//The order from Siemens is complete, nothing is remembered from earlier washes.
//Local requests of FB_CIP_Siemens carry their start too, requests of the HMI have none (item 7, 02.11.2026)
IF eReq.eClient=E_CIP_Usage.eExternal OR eReq.eStartState<>E_Element_State_Long.eOff THEN;
	eCIP_State:=eReq.eStartState;
ELSIF eReq.eType=E_CIP_Type.Full THEN;
	eCIP_State:=E_Element_State_Long.eNotClean;
ELSE;
	eCIP_State:=E_Element_State_Long.eCIP_1_Rinzed;
END_IF
g_Data.b_CIP_Run:=TRUE;
bClientRef_done:=TRUE;
END_ACTION

ACTION _aReadyToCondition_Count_active:

(*
IF TRUE 
AND pcFlow1_Rate.mRun()
AND pcFlow2_Rate.mRun()
//AND pcPressure.mRun()
THEN;
	bStepDone:=TRUE;
ELSE;
	bStepDone:=FALSE;
END_IF
*)
END_ACTION

ACTION _aReadyToCondition_Count_entry:

fb_PumpCIP.m_Run(RPM:=st_CIP_Param.r_CIP_Pump);
END_ACTION

ACTION _aReFill_Water_T93_active:
IF TRUE
//AND lvlTank_T94.e_state=E_Tank_Level.eLL
AND lvlTank_T93.rTankLevel + 0 > st_CIP_Param.r_Tank93_Volume//st_CIP_Param.r_Water_TankLvl_Lcl_1 // Client requered Level
THEN;	
	bStepDone:=TRUE;
	fbPis.m_SetByRecipe(stPis:=stPis_FillWater_T93, req:=E_Piston_Recipe_State.Release);
ELSE;
	//Fill water
	bStepDone:=FALSE;
		IF NOT arrTanksSens[E_Tank_Name.T93].get_stTankLevel_OverFlow() THEN;
			fbPis.m_SetByRecipe(stPis:=stPis_FillWater_T93, req:=E_Piston_Recipe_State.Act);			
		END_IF
END_IF
END_ACTION

ACTION _aReFill_Water_T94_active:
IF TRUE
//AND lvlTank_T94.e_state=E_Tank_Level.eLL
AND lvlTank_T94.rTankLevel +20>st_CIP_Param.r_Tank94_Volume//st_CIP_Param.r_Water_TankLvl_Lcl_1 // Client requered Level
THEN;	
	bStepDone:=TRUE;
	fbPis.m_SetByRecipe(stPis:=stPis_FillWater_T94, req:=E_Piston_Recipe_State.Release);
ELSE;
	//Fill water
	bStepDone:=FALSE;
	IF NOT arrTanksSens[E_Tank_Name.T94].get_stTankLevel_OverFlow() THEN;
		fbPis.m_SetByRecipe(stPis:=stPis_FillWater_T94, req:=E_Piston_Recipe_State.Act);			
	END_IF
END_IF
END_ACTION

ACTION _aReset_Cond_Tm_CIP2_01_active:
tonr_CIP_Condition(ResetTime:=TRUE);
END_ACTION

ACTION _aSet_Valves_ToDeafult_active:
bStepDone:=FALSE;
IF TRUE 
AND fbPis.m_CheckByRecipe(stPis:=stPis_FillWater_T91, 	req:=E_Piston_Recipe_State.Release) 
AND fbPis.m_CheckByRecipe(stPis:=stPis_FillWater_T92, 	req:=E_Piston_Recipe_State.Release) 
AND fbPis.m_CheckByRecipe(stPis:=stPis_FillWater_T93, 	req:=E_Piston_Recipe_State.Release) 
AND fbPis.m_CheckByRecipe(stPis:=stPis_FillWater_T94, 	req:=E_Piston_Recipe_State.Release) 

THEN;
	bStepDone:=TRUE;
END_IF
END_ACTION

ACTION _aSet_Valves_ToDeafult_entry:
fbPis.m_SetByRecipe(stPis:=stPis_FillWater_T91, req:=E_Piston_Recipe_State.Release);
fbPis.m_SetByRecipe(stPis:=stPis_FillWater_T92, req:=E_Piston_Recipe_State.Release);
fbPis.m_SetByRecipe(stPis:=stPis_FillWater_T93, req:=E_Piston_Recipe_State.Release);
fbPis.m_SetByRecipe(stPis:=stPis_FillWater_T94, req:=E_Piston_Recipe_State.Release);

_aDisconnect_n_Drain_CIP_Client_entry();
END_ACTION

ACTION _aSprinkler_Request_CIP1_active:


IF TRUE // Type Tank
AND bClientTypeIs_Tank	
AND bSprinkler
THEN;	
	bStepDone:=TRUE;
	m_DashState_done(stage:=E_CIP_DashStage_List.e02_CIP1_Client_Drain_Product_Rest_Sprinkler);
	
ELSIF TRUE // Type Pine
AND NOT bClientTypeIs_Tank	
THEN;	
	bStepDone:=TRUE;
	m_DashState_done(stage:=E_CIP_DashStage_List.e01_CIP1_Client_Drain_Product_Rest_Pipe);
	
ELSE;
	//continue with sprinkler
	bStepDone:=FALSE;
	m_DashState_done(stage:=E_CIP_DashStage_List.e01_CIP1_Client_Drain_Product_Rest_Pipe);
	m_DashState_activate(stage:=E_CIP_DashStage_List.e02_CIP1_Client_Drain_Product_Rest_Sprinkler);
	
END_IF
END_ACTION

ACTION _aSprinkler_Request_CIP35_active:


IF TRUE // Type Tank
AND bClientTypeIs_Tank	
AND bSprinkler
THEN;	
	bStepDone:=TRUE;
	CASE eCIP_State OF
	
		E_Element_State_Long.eCIP_2_Deterged:;
				m_DashState_done(stage:=E_CIP_DashStage_List.e11_CIP3_Detergent_Clean_Sprinkler);
	
		E_Element_State_Long.eCIP_4_Sanitized:;
				m_DashState_done(stage:=E_CIP_DashStage_List.e20_CIP5_DisInfection_Clean_Sprinkler);
				
	END_CASE	
	
ELSIF TRUE // Type Pine
AND NOT bClientTypeIs_Tank	
THEN;	
	bStepDone:=TRUE;
	CASE eCIP_State OF
	
		E_Element_State_Long.eCIP_2_Deterged:;
				m_DashState_done(stage:=E_CIP_DashStage_List.e10_CIP3_Detergent_Clean_Pipe);
	
		E_Element_State_Long.eCIP_4_Sanitized:;
				m_DashState_done(stage:=E_CIP_DashStage_List.e19_CIP5_DisInfection_Clean_Pipe);
				
	END_CASE	
	
ELSE;
	//continue with sprinkler
	bStepDone:=FALSE;
	CASE eCIP_State OF
	
		E_Element_State_Long.eCIP_2_Deterged:;
				m_DashState_done(stage:=E_CIP_DashStage_List.e10_CIP3_Detergent_Clean_Pipe);
				m_DashState_activate(stage:=E_CIP_DashStage_List.e11_CIP3_Detergent_Clean_Sprinkler);
	
		E_Element_State_Long.eCIP_4_Sanitized:;
				m_DashState_done(stage:=E_CIP_DashStage_List.e19_CIP5_DisInfection_Clean_Pipe);
				m_DashState_activate(stage:=E_CIP_DashStage_List.e20_CIP5_DisInfection_Clean_Sprinkler);
				
	END_CASE	
	
END_IF
END_ACTION

ACTION _aStartPump_CIP1_01_active:
bStepDone:=FALSE;
(*
IF StartPump_CIP1_01.t>SECOND_TO_TIME(st_CIP_Param.t_PumpInitRun) 
OR lvlTank_T93.rTankLevel<st_CIP_Param.r_Tank93_Volume//st_CIP_Param.r_RWater_93_TankLvl
THEN//Time+flow+water volume
	bStepDone:=TRUE;
END_IF
*)
bStepDone:=TRUE;
END_ACTION

ACTION _aStartPump_CIP1_01_entry:
fb_PumpCIP.m_Run(RPM:=st_CIP_Param.r_CIP_Pump);


mVolumeReset_All();

tonr_CIP_Condition(ResetTime:=TRUE);
END_ACTION

ACTION _aStartPump_CIP2_01_active:
IF TRUE 
//AND stAnalogSensor[E_ASense_Name.FT1001].Value>=g_Data.arr_CIP_Recipe[0].r_Flow_1 // 
//AND stAnalogSensor[E_ASense_Name.FT1002].Value>=g_Data.arr_CIP_Recipe[0].r_Flow_2 // 
//AND stAnalogSensor[E_ASense_Name.PT1001].Value>=g_Data.arr_CIP_Recipe[0].r_Pressure // 
//AND pcFlow1_Rate.mRun_With_SP(Set_Point:=g_Data.arr_CIP_Recipe[0].r_Flow_Pipe)
//AND pcFlow2_Rate.mRun_With_SP(Set_Point:=g_Data.arr_CIP_Recipe[0].r_Flow_Pipe)
AND pcFlow1_Rate.mRun()
AND pcFlow2_Rate.mRun()
//AND pcPressure.mRun()
THEN;
	bStepDone:=TRUE;
ELSE;
	bStepDone:=FALSE;
END_IF

fb_PumpCIP.m_Run(RPM:=pcFlow1_Rate.mRun_PID(Set_Point:=g_Data.arr_CIP_Recipe[0].r_Flow_Pipe,controlManual:=NOT(fb_PumpCIP.modeAuto)));
END_ACTION

ACTION _aStartPump_CIP2_01_entry:

//fb_PumpDetergent.m_Auto();
fb_HeatExchenger.m_Auto();
bCIP_Condition_Failed:=FALSE;
bCIP_Condition_Done:=FALSE;
iConcentrationDeluteCounter:=0;

nStepHeat:=1;
END_ACTION

ACTION _aStartPump_CIP2_02_active:
fb_PumpCIP.m_Run(RPM:=pcFlow1_Rate.mRun_PID(Set_Point:=fFlowRate, controlManual:=NOT(fb_PumpCIP.modeAuto)));


IF TRUE 
AND pcFlow1_Rate.mRun()
AND pcFlow2_Rate.mRun()
//AND pcPressure.mRun()
THEN;
	bStepDone:=TRUE;
ELSE;
	bStepDone:=FALSE;
END_IF
END_ACTION

ACTION _aStartPump_CIP2_02_entry:
fb_HeatExchenger.m_Auto();
bCIP_Condition_Failed:=FALSE;
bCIP_Condition_Done:=FALSE;
iConcentrationDeluteCounter:=0;

nStepHeat:=10;
END_ACTION

ACTION _aStartPump_CIP2_RPM_01_active:
bStepDone:=FALSE;
fb_PumpCIP.m_Run(RPM:=g_Data.arr_CIP_Recipe[0].r_CIP_Pump);//1500

IF TRUE //Future condition
AND StartPump_CIP2_RPM_01.t>SECOND_TO_TIME(g_Data.arr_CIP_Recipe[0].t_PumpInitRun) 
AND fb_PumpCIP.nRPM=g_Data.arr_CIP_Recipe[0].r_CIP_Pump
//AND stAnalogSensor[E_ASense_Name.FT1001].Value>=g_Data.arr_CIP_Recipe[0].r_Flow_Pipe // 
//AND stAnalogSensor[E_ASense_Name.FT1002].Value>=g_Data.arr_CIP_Recipe[0].r_Flow_Pipe // 
THEN;
	bStepDone:=TRUE;
END_IF
END_ACTION

ACTION _aStartPump_CIP2_RPM_02_active:
bStepDone:=FALSE;

fb_PumpCIP.m_Run(RPM:=st_CIP_Param.r_CIP_Pump);

bStepDone:=TRUE;

// to stas question ? deference:
//fb_PumpCIP.m_Run(RPM:=g_Data.arr_CIP_Recipe[0].r_CIP_Pmp_1);//1500
//fb_PumpCIP.m_Run(RPM:=st_CIP_Param.r_CIP_Pmp_1);
(*
IF TRUE //Future condition
AND delta_T92_Volume < - st_CIP_Param.r_Volume_Solution_Fill // Volume 
//AND StartPump_CIP2_RPM_02.t>SECOND_TO_TIME(g_Data.arr_CIP_Recipe[0].t_PumpInitRun) 
THEN;
	bStepDone:=TRUE;
END_IF
*)
END_ACTION

ACTION _aStartPump_CIP2_RPM_02_entry:
mVolumeReset_All();
tonr_CIP_Condition(ResetTime:=TRUE);
END_ACTION

ACTION _aStartPump_CIP4_RPM_01_active:
bStepDone:=FALSE;
fb_PumpCIP.m_Run(RPM:=g_Data.arr_CIP_Recipe[0].r_CIP_Pump);

IF TRUE //Future condition
AND StartPump_CIP4_RPM_01.t>SECOND_TO_TIME(g_Data.arr_CIP_Recipe[0].t_PumpInitRun) 
THEN;
	bStepDone:=TRUE;
END_IF
END_ACTION

ACTION _aStartPump_CIP4_RPM_02_active:
bStepDone:=FALSE;
fb_PumpCIP.m_Run(RPM:=pcFlow1_Rate.mRun_PID(Set_Point:=st_CIP_Param.r_CIP_Pump,controlManual:=NOT(fb_PumpCIP.modeAuto)));


IF TRUE //Future condition
AND StartPump_CIP4_RPM_02.t>SECOND_TO_TIME(st_CIP_Param.t_PumpInitRun) 
THEN;
	bStepDone:=TRUE;
END_IF
END_ACTION

ACTION _aStartPump_CIP4_01_active:
IF TRUE 
(*AND stAnalogSensor[E_ASense_Name.FT1001].Value>=g_Data.arr_CIP_Recipe[0].r_Flow_1//200 // 
AND stAnalogSensor[E_ASense_Name.FT1002].Value>=g_Data.arr_CIP_Recipe[0].r_Flow_2//200 // 
AND stAnalogSensor[E_ASense_Name.PT1001].Value>=g_Data.arr_CIP_Recipe[0].r_Pressure//0.5 //*)
AND pcFlow1_Rate.mRun()
AND pcFlow2_Rate.mRun()
//AND pcPressure.mRun()
THEN;
	bStepDone:=TRUE;
ELSE;
	bStepDone:=FALSE;
END_IF

fb_PumpCIP.m_Run(RPM:=pcFlow1_Rate.mRun_PID(Set_Point:=g_Data.arr_CIP_Recipe[0].r_Flow_Pipe,controlManual:=NOT(fb_PumpCIP.modeAuto)));
END_ACTION

ACTION _aStartPump_CIP4_01_entry:


fb_HeatExchenger.m_Auto();
bCIP_Condition_Failed:=FALSE;
bCIP_Condition_Done:=FALSE;

nStepHeat:=2;
iConcentrationDeluteCounter:=0;
END_ACTION

ACTION _aStartPump_CIP4_02_active:
IF TRUE 
(*AND stAnalogSensor[E_ASense_Name.FT1001].Value>=st_CIP_Param.r_Flow_1 // 
AND stAnalogSensor[E_ASense_Name.FT1002].Value>=st_CIP_Param.r_Flow_2 // 
AND stAnalogSensor[E_ASense_Name.PT1001].Value>=st_CIP_Param.r_Pressure // *)
AND pcFlow1_Rate.mRun()
AND pcFlow2_Rate.mRun()
//AND pcPressure.mRun()
THEN;
	bStepDone:=TRUE;
ELSE;
	bStepDone:=FALSE;
END_IF

//fb_PumpCIP.m_Run(RPM:=pcFlow1_Rate.mRun_PID(Set_Point:=fFlowRate,controlManual:=NOT(fb_PumpCIP.modeAuto)));

IF TRUE //Future condition
AND StartPump_CIP4_02.t>SECOND_TO_TIME(st_CIP_Param.t_PumpInitRun) THEN;
	fb_PumpCIP.m_Run(RPM:=pcFlow1_Rate.mRun_PID(Set_Point:=fFlowRate,controlManual:=NOT(fb_PumpCIP.modeAuto)));
	
END_IF

IF NOT bSprinkler THEN
	//pipe
	tConditionTime	:=st_CIP_Param.t_ConditionDisInfection;
	fFlowRate		:=st_CIP_Param.r_Flow_Pipe;
	//rVolume_Collect :=st_CIP_Param.r_Volume_Collect_DisInfection;
	//rVolume_Drain	:=st_CIP_Param.r_Volume_Drain_DisInfection;
	//rVolume_Recycle	:=st_CIP_Param.r_Volume_Recycle_DisInfection;
ELSE
	//sprinkler
	tConditionTime	:=st_CIP_Param.t_ConditionDisInfection_Sprinkler;
	fFlowRate		:=st_CIP_Param.r_Flow_Sprinkler;
	//rVolume_Collect :=st_CIP_Param.r_Volume_Collect_DisInfection*st_CIP_Param.r_Volume_Sprinkler_Ratio;
	//rVolume_Drain	:=st_CIP_Param.r_Volume_Drain_DisInfection*st_CIP_Param.r_Volume_Sprinkler_Ratio;
	//rVolume_Recycle	:=st_CIP_Param.r_Volume_Recycle_DisInfection*st_CIP_Param.r_Volume_Sprinkler_Ratio;
END_IF
END_ACTION

ACTION _aStartPump_CIP4_02_entry:

//fb_PumpDisinfection.m_Auto();
	
//Heat Exchenger	
fb_HeatExchenger.m_Auto();

bCIP_Condition_Failed:=FALSE;
bCIP_Condition_Done:=FALSE;
iConcentrationDeluteCounter:=0;

nStepHeat:=20;
END_ACTION

ACTION _aStartPump_CIP35_active:
bStepDone:=FALSE;
IF TRUE 
//AND fbPis.m_CheckByRecipe(stPis:=stPis_FillWater_T94, 		req:=E_Piston_Recipe_State.NoChanges) 
THEN
	//bStepDone:=TRUE;
END_IF
bStepDone:=TRUE;
END_ACTION

ACTION _aStartPump_CIP35_entry:
//fbPis.m_SetByRecipe(stPis:=stPis_FillWater_T94, 	req:=E_Piston_Recipe_State.NoChanges);
fb_PumpCIP.m_Run(RPM:=st_CIP_Param.r_CIP_Pump);


mVolumeReset_All();
bSprinkler:=FALSE;
tonr_CIP_Condition(ResetTime:=TRUE);
END_ACTION

ACTION _aStop_Pump_entry:
fb_PumpCIP.m_Stop();


fb_PumpDetergent.m_Stop();
fb_PumpDisinfection.m_Stop();
END_ACTION

ACTION _aStopPump_CIP1_01_entry:
fb_PumpCIP.m_Stop();
END_ACTION

ACTION _aStopPump_CIP1_02_entry:
fb_PumpCIP.m_Stop();
END_ACTION

ACTION _aStopPump_CIP2_01_entry:
fb_PumpCIP.m_Stop();

m_DashState_done(stage:=E_CIP_DashStage_List.e04_CIP2_Local_Detergent_Condition);
END_ACTION

ACTION _aStopPump_CIP2_02_entry:
fb_PumpCIP.m_Stop();
END_ACTION

ACTION _aStopPump_CIP2_03_entry:
fb_PumpCIP.m_Stop();
END_ACTION

ACTION _aStopPump_CIP4_01_entry:
fb_PumpCIP.m_Stop();

m_DashState_done(stage:=E_CIP_DashStage_List.e13_CIP4_Local_DisInfection_Condition);
END_ACTION

ACTION _aStopPump_CIP4_02_entry:
fb_PumpCIP.m_Stop();
END_ACTION

ACTION _aStopPump_CIP4_03_entry:
fb_PumpCIP.m_Stop();
END_ACTION

ACTION _aStopPump_CIP35_01_entry:
fb_PumpCIP.m_Stop();
END_ACTION

ACTION _aStopPump_CIP35_02_entry:
fb_PumpCIP.m_Stop();
END_ACTION

ACTION _aTank_LowLevel_CIP1_01_active:
bStepDone:=m_Check_ProductionTank_Low_Level();
END_ACTION

ACTION _aTank_LowLevel_CIP1_02_active:
bStepDone:=m_Check_ProductionTank_Low_Level();
END_ACTION

ACTION _aTank_LowLevel_CIP1_02_entry:
fb_PumpCIP.m_Stop();
END_ACTION

ACTION _aTank_LowLevel_CIP2_01_active:
bStepDone:=m_Check_ProductionTank_Low_Level();
END_ACTION

ACTION _aTank_LowLevel_CIP2_02_active:
bStepDone:=m_Check_ProductionTank_Low_Level();
END_ACTION

ACTION _aTank_LowLevel_CIP2_02_entry:
fb_PumpCIP.m_Stop();
END_ACTION

ACTION _aTank_LowLevel_CIP4_01_active:
bStepDone:=m_Check_ProductionTank_Low_Level();
END_ACTION

ACTION _aTank_LowLevel_CIP4_02_active:
bStepDone:=m_Check_ProductionTank_Low_Level();
END_ACTION

ACTION _aTank_LowLevel_CIP4_02_entry:
fb_PumpCIP.m_Stop();
END_ACTION

ACTION _aTank_LowLevel_CIP35_01_active:
bStepDone:=m_Check_ProductionTank_Low_Level();
END_ACTION

ACTION _aTank_LowLevel_CIP35_02_active:
bStepDone:=m_Check_ProductionTank_Low_Level();
END_ACTION

ACTION _aTank_LowLevel_CIP35_02_entry:
fb_PumpCIP.m_Stop();
END_ACTION

ACTION _aTank_MixProof_Clean_CIP2_active:
//Mix-proof valves are on the plant side
bStepDone:=TRUE;
END_ACTION

ACTION _aTank_MixProof_Clean_CIP2_entry:
fb_PumpCIP.m_Stop();
END_ACTION

ACTION _aTank_MixProof_Clean_CIP4_active:
//Mix-proof valves are on the plant side
bStepDone:=TRUE;
END_ACTION

ACTION _aTank_MixProof_Clean_CIP4_entry:
fb_PumpCIP.m_Stop();
END_ACTION

ACTION _aTriBlender_Selection_active:
bStepDone:=TRUE;
END_ACTION

ACTION _aTriBlender_Selection_entry:

END_ACTION

ACTION _aWaiting_Client_Drain_Done_active:
// The command from Set_Valves_ToDeafult is lost if a sub-FB was in Init or busy: give it again
IF fbCIP_Source.m_IsFree() AND NOT fbCIP_Source.m_CheckStatus(eReqStatus:=E_CIP_Source.eClose) THEN;
	fbCIP_Source.m_Run(eReqProc:=E_CIP_Source.eClose);
END_IF
IF fbCIP_Usage.m_IsFree() AND NOT fbCIP_Usage.m_CheckStatus(eReqStatus:=E_CIP_Usage.eLocal) THEN;
	fbCIP_Usage.m_Run(eReqProc:=E_CIP_Usage.eLocal);
END_IF
IF fbCIP_Return.m_IsFree() AND NOT fbCIP_Return.m_CheckStatus(eReqStatus:=E_CIP_Return.eDrain) THEN;
	fbCIP_Return.m_Run(eReqProc:=E_CIP_Return.eDrain);
END_IF

_aDisconnect_n_Drain_CIP_Client_active();
END_ACTION

ACTION act_CallProcessControl:
//Heat Exchanger
	stHeatExchanger.rValue:=g_AnalogSensor.stAnalogSensor[E_ASense_Name.TT1105].Value;
	//stHeatExchanger.rSetPoint:=st_CIP_Param.r_Temper_ClientReturn;
	pcHeatExchanger(stProcessControl:=stHeatExchanger );
//Client temperature return
	stTemp_ClntReturn.rValue:=g_AnalogSensor.stAnalogSensor[E_ASense_Name.TT1101].Value;//gIO.fbScaleFactor[E_ASense_Name.TT1101].rValOut;
	//stTemp_ClntReturn.rSetPoint:=st_CIP_Param.n _ClientReturn;
	pcTemp_ClntReturn(stProcessControl:=stTemp_ClntReturn );

//Detergent
	//Concentration
	stDetergent.rValue:=g_AnalogSensor.stAnalogSensor[E_ASense_Name.CT1101_3].Value;
	//###stDetergent.ToleranceHigh:=0.05;
	//###stDetergent.ToleravceLow:=0.05;
	//###stDetergent.rSetPoint:=st_CIP_Param.r_DetergentConcentration;//0.3;
	pcDetergent(stProcessControl:=stDetergent );
		
	//Temperature
	//stTemperature_Deterg.rValue:=testTemperature;
	stTemperature_Deterg.rValue:=g_AnalogSensor.stAnalogSensor[E_ASense_Name.TT1003].Value;
	//###stTemperature_Deterg.ToleranceHigh:=1;
	//###stTemperature_Deterg.ToleravceLow:=1;
	//###stTemperature_Deterg.rSetPoint:=st_CIP_Param.r_Temper_Detergent;
	pcTemperature_Deterg(stProcessControl:=stTemperature_Deterg );


//Disinfectant
	//Concentration
	stDisInfectant.rValue:=g_AnalogSensor.stAnalogSensor[E_ASense_Name.CT1101_4].Value;
	//###stDisInfectant.ToleranceHigh:=0.05;
	//###stDisInfectant.ToleravceLow:=0.05;
	//###stDisInfectant.rSetPoint:=st_CIP_Param.r_DisInfectionConcentration;//0.3;
	pcDisInfectant(stProcessControl:=stDisInfectant );
		
	//Temperature	
	//stTemperature_Dis.rValue:=testTemperature;
	stTemperature_Dis.rValue:=g_AnalogSensor.stAnalogSensor[E_ASense_Name.TT1004].Value;
	//###stTemperature_Dis.ToleranceHigh:=1;//0.5
	//###stTemperature_Dis.ToleravceLow:=1;//0.5
	//###stTemperature_Dis.rSetPoint:=st_CIP_Param.r_Temper_DisInfection;//65;
	pcTemperature_Dis(stProcessControl:=stTemperature_Dis );	
	
// Flow_Rate
	//CIP Pump
		//Pump CIP infeed
		stFlow1_Rate.rValue:=g_AnalogSensor.stAnalogSensor[E_ASense_Name.FT1001].Value;
		stFlow1_Rate.rValue:=g_AnalogSensor.stAnalogSensor[E_ASense_Name.FT1001].Value;
		stFlow1_Rate.rValue_Min_To_ReleaseControl:=50;// Litter/Hours
		//stFlow1_Rate.rSetPoint:=st_CIP_Param.r_Flow_Pipe;//:=150
		stFlow1_Rate.bPause:=stOper[E_ModeZone.eCIP].iActOperation=E_OperationButtons.ePauseAll;
		stFlow1_Rate.fCtrlOutput_Manual:=fb_PumpCIP.nRPM;
		stFlow1_Rate.fCtrlOutput_Max:=1700;
		stFlow1_Rate.fCtrlOutput_Min:=700;
		pcFlow1_Rate(stProcessControl:=stFlow1_Rate, );

		//Pump CIP return 
		stFlow2_Rate.rValue:=g_AnalogSensor.stAnalogSensor[E_ASense_Name.FT1002].Value;
		stFlow3_Rate.rValue:=g_AnalogSensor.stAnalogSensor[E_ASense_Name.FT1002].Value;
		stFlow3_Rate.rSetPoint:=stFlow2_Rate.rSetPoint;
		pcFlow2_Rate(stProcessControl:=stFlow2_Rate );
		pcFlow3_Rate(stProcessControl:=stFlow3_Rate );

		// TBD : to check if the first loop(local prepare) when Client selected gets relevant Flow SetPoint 
		IF bSprinkler THEN
			stFlow1_Rate.rSetPoint:=st_CIP_Param.r_Flow_Sprinkler;
			stFlow2_Rate.rSetPoint:=st_CIP_Param.r_Flow_Sprinkler;
		ELSE
			stFlow1_Rate.rSetPoint:=st_CIP_Param.r_Flow_Pipe;
			stFlow2_Rate.rSetPoint:=st_CIP_Param.r_Flow_Pipe;
		END_IF		
		
	//CIP Client Color pump
		//stFlow_Rate.rSetPoint:=150;
	//CIP Client Marinada pump
		//stFlow_Rate.rSetPoint:=150;
		
//Presure
		stP1001_Pressure.rValue:=g_AnalogSensor.stAnalogSensor[E_ASense_Name.PT1001].Value;
		pcP1001_Pressure(stProcessControl:=stP1001_Pressure );


//Load def set points
IF bLoadDefSetPoints THEN
	bLoadDefSetPoints:=FALSE;
	mLoadDefProcessSetPoints();
END_IF
		
//selecting set point based on user
	
	IF bTestPID THEN;
		pcFlow1_Rate.mRun();

		fb_PumpCIP.m_Auto(control:=pcFlow1_Rate.mRun_PID(Set_Point:=180,controlManual:=NOT(fb_PumpCIP.modeAuto)));
		
		//by CIP Pump RPM control		
		
		IF fb_PumpCIP.modeAuto THEN;
			stFlow1_Rate.bManual:=FALSE;
		ELSE;
			stFlow1_Rate.bManual:=TRUE;
			stFlow1_Rate.fCtrlOutput_Manual:=fb_PumpCIP.nRPM;
		END_IF
		
			
	END_IF
END_ACTION

ACTION act_GetReference:
stPis_FillWater_T91 REF= stPis[valFillWater_T91];
stPis_FillWater_T92 REF= stPis[valFillWater_T92];
stPis_FillWater_T93 REF= stPis[valFillWater_T93];
stPis_FillWater_T94 REF= stPis[valFillWater_T94];

	//concentration
stDetergent 	REF=g_ProcControl.arr_stProcCntrl[E_ProcessControl_Name.eDetergentConc];
pcDetergent 	REF=g_ProcControl.arr_fbProcCntrl[E_ProcessControl_Name.eDetergentConc];

stDisInfectant 	REF=g_ProcControl.arr_stProcCntrl[E_ProcessControl_Name.eDisinfectionConc];
pcDisInfectant 	REF=g_ProcControl.arr_fbProcCntrl[E_ProcessControl_Name.eDisinfectionConc];

	//Temperature
stTemperature_Deterg REF=g_ProcControl.arr_stProcCntrl[E_ProcessControl_Name.eDeterTemp];
pcTemperature_Deterg REF=g_ProcControl.arr_fbProcCntrl[E_ProcessControl_Name.eDeterTemp];

stTemperature_Dis 	 REF=g_ProcControl.arr_stProcCntrl[E_ProcessControl_Name.eDisTemp];
pcTemperature_Dis 	 REF=g_ProcControl.arr_fbProcCntrl[E_ProcessControl_Name.eDisTemp];
	//Flow rate
stFlow1_Rate REF=g_ProcControl.arr_stProcCntrl[E_ProcessControl_Name.eCIP_Flow_1];
pcFlow1_Rate REF=g_ProcControl.arr_fbProcCntrl[E_ProcessControl_Name.eCIP_Flow_1];

stFlow2_Rate REF=g_ProcControl.arr_stProcCntrl[E_ProcessControl_Name.eCIP_Flow_2];
pcFlow2_Rate REF=g_ProcControl.arr_fbProcCntrl[E_ProcessControl_Name.eCIP_Flow_2];

stFlow3_Rate REF=g_ProcControl.arr_stProcCntrl[E_ProcessControl_Name.eCIP_Flow_3];
pcFlow3_Rate REF=g_ProcControl.arr_fbProcCntrl[E_ProcessControl_Name.eCIP_Flow_3];

	//Level

	//Pressure
stP1001_Pressure 	REF=g_ProcControl.arr_stProcCntrl[E_ProcessControl_Name.eCIP_Pressure];
pcP1001_Pressure 	REF=g_ProcControl.arr_fbProcCntrl[E_ProcessControl_Name.eCIP_Pressure];

//temperature control
stTemp_ClntReturn REF=g_ProcControl.arr_stProcCntrl[E_ProcessControl_Name.eClientReturn_Temp];
pcTemp_ClntReturn REF=g_ProcControl.arr_fbProcCntrl[E_ProcessControl_Name.eClientReturn_Temp];

stHeatExchanger REF=g_ProcControl.arr_stProcCntrl[E_ProcessControl_Name.eHeatExchanger];
pcHeatExchanger REF=g_ProcControl.arr_fbProcCntrl[E_ProcessControl_Name.eHeatExchanger];
END_ACTION

ACTION act_HeatExchng:
//calling heat exchanger 
fb_HeatExchenger(stHeatExchanger:=g_Data.stHeatExchanger );

//Choosing heat exchanger set point 

CASE nStepHeat OF
	0:	
	(*	//heat excahnger not in use 
	1:
		//detergent local
		IF stTemperature_Deterg.Control_ON THEN
			g_Data.stHeatExchanger:=stTemperature_Deterg.Control_Value;
		ELSE
			g_Data.stHeatExchanger:=0;
		END_IF
	10:
		//detergent client
	2:
		//disinfection
		IF stTemperature_Dis.Control_ON THEN
			g_Data.stHeatExchanger:=stTemperature_Dis.Control_Value;
		ELSE
			g_Data.stHeatExchanger:=0;
		END_IF
	20:
		//disinfection client
	3:
		//something else
		*)
END_CASE
END_ACTION

ACTION act_Oper:
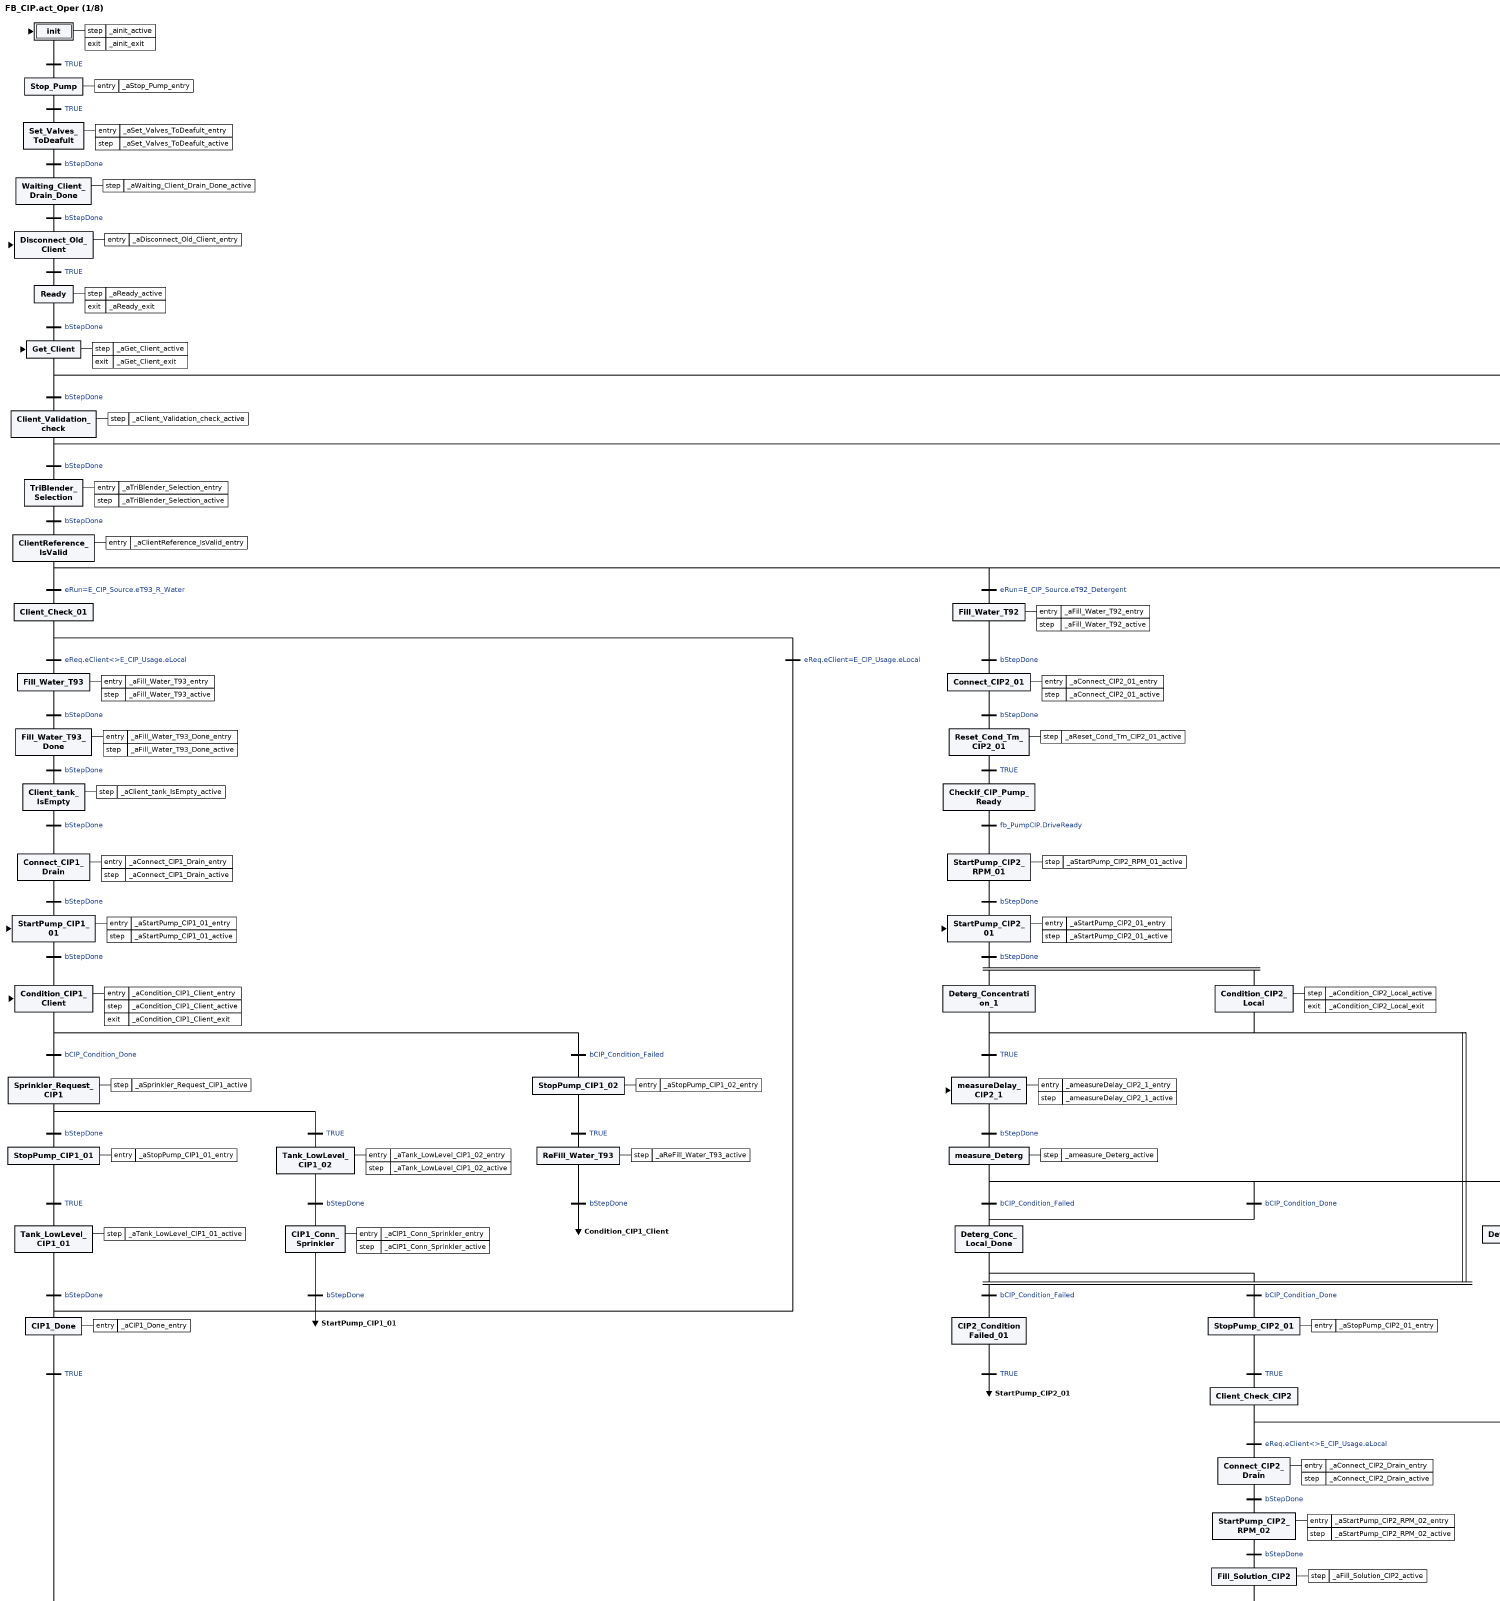
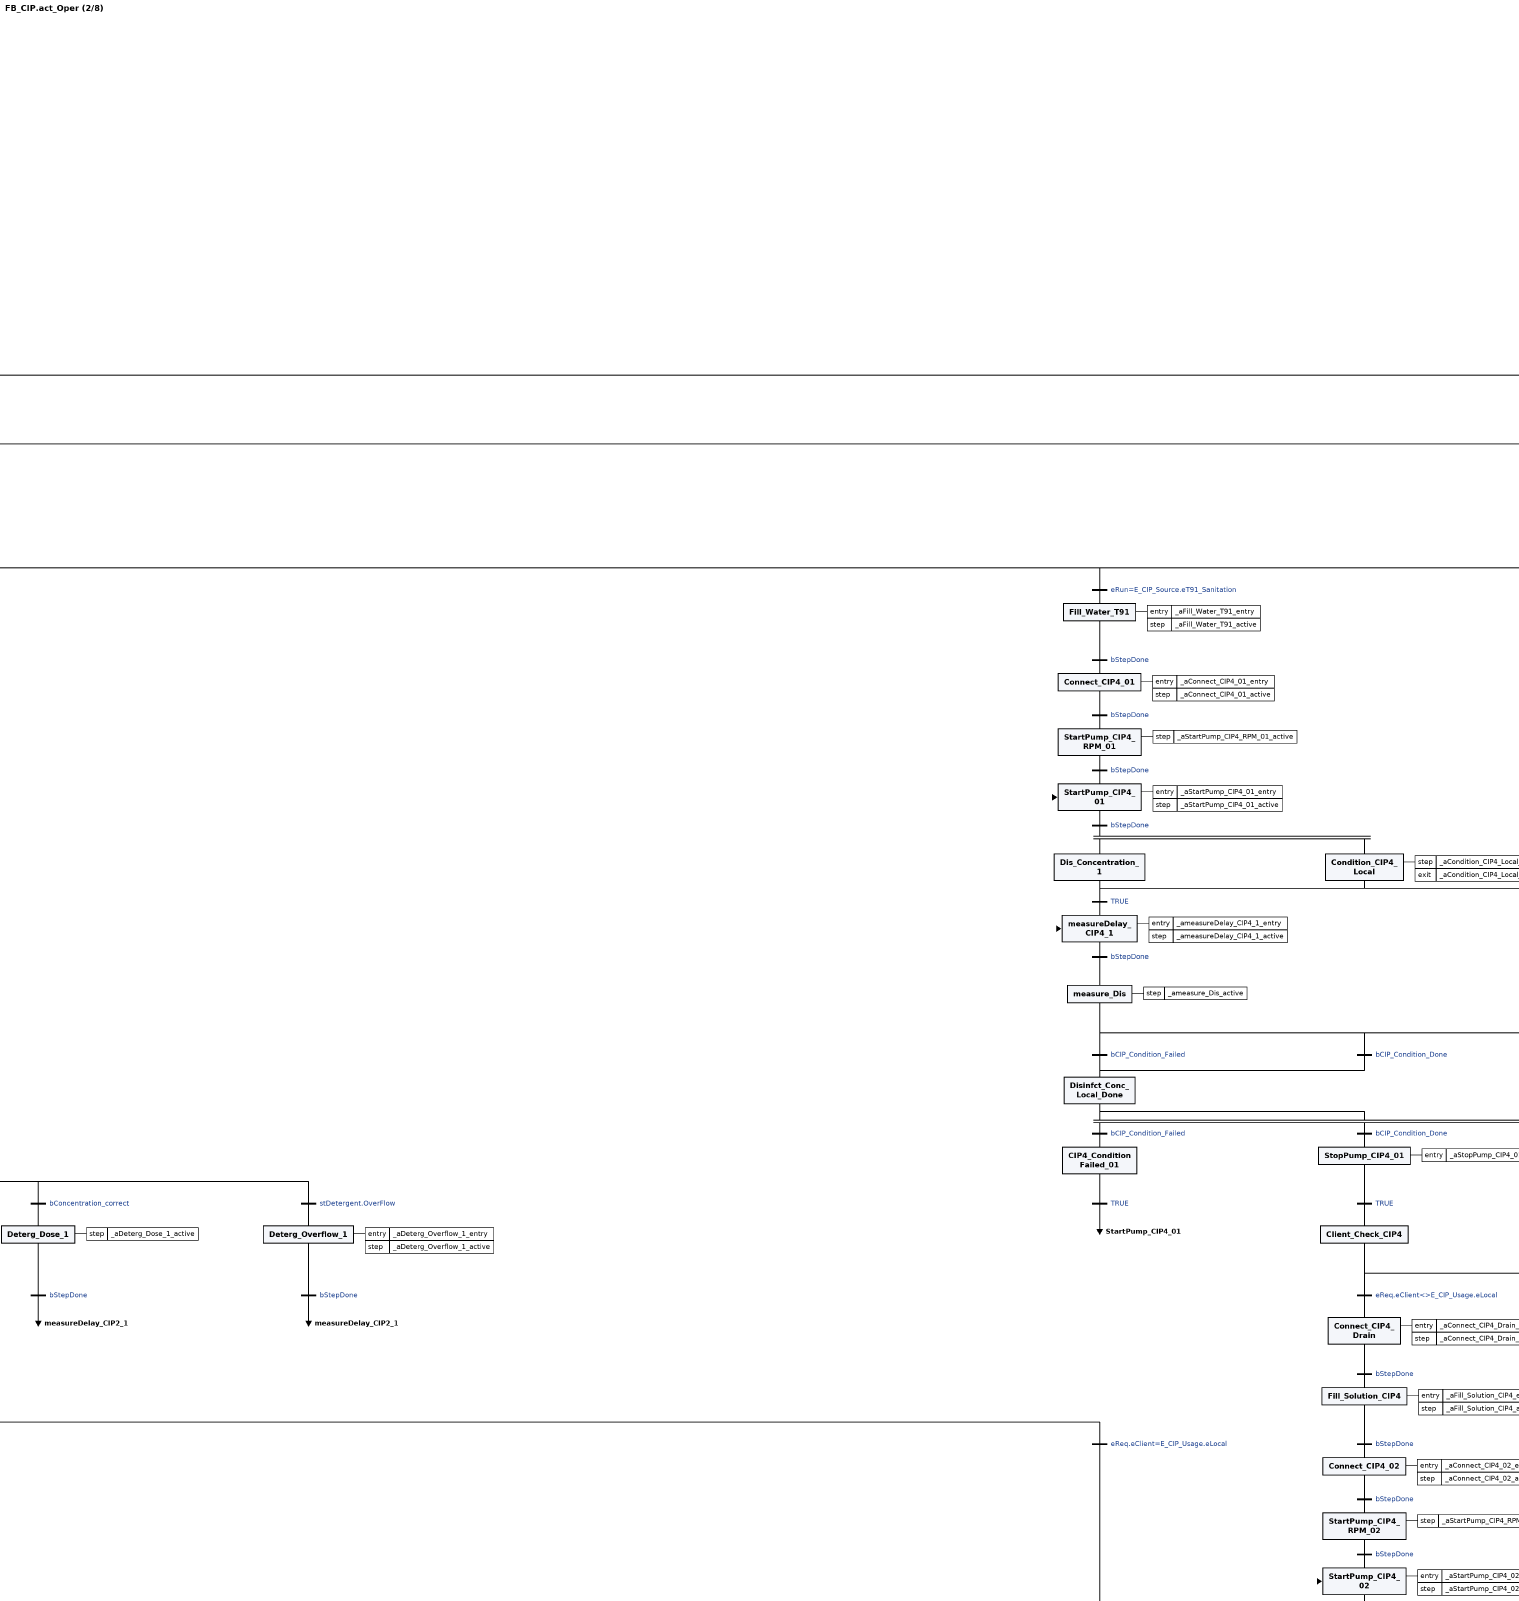
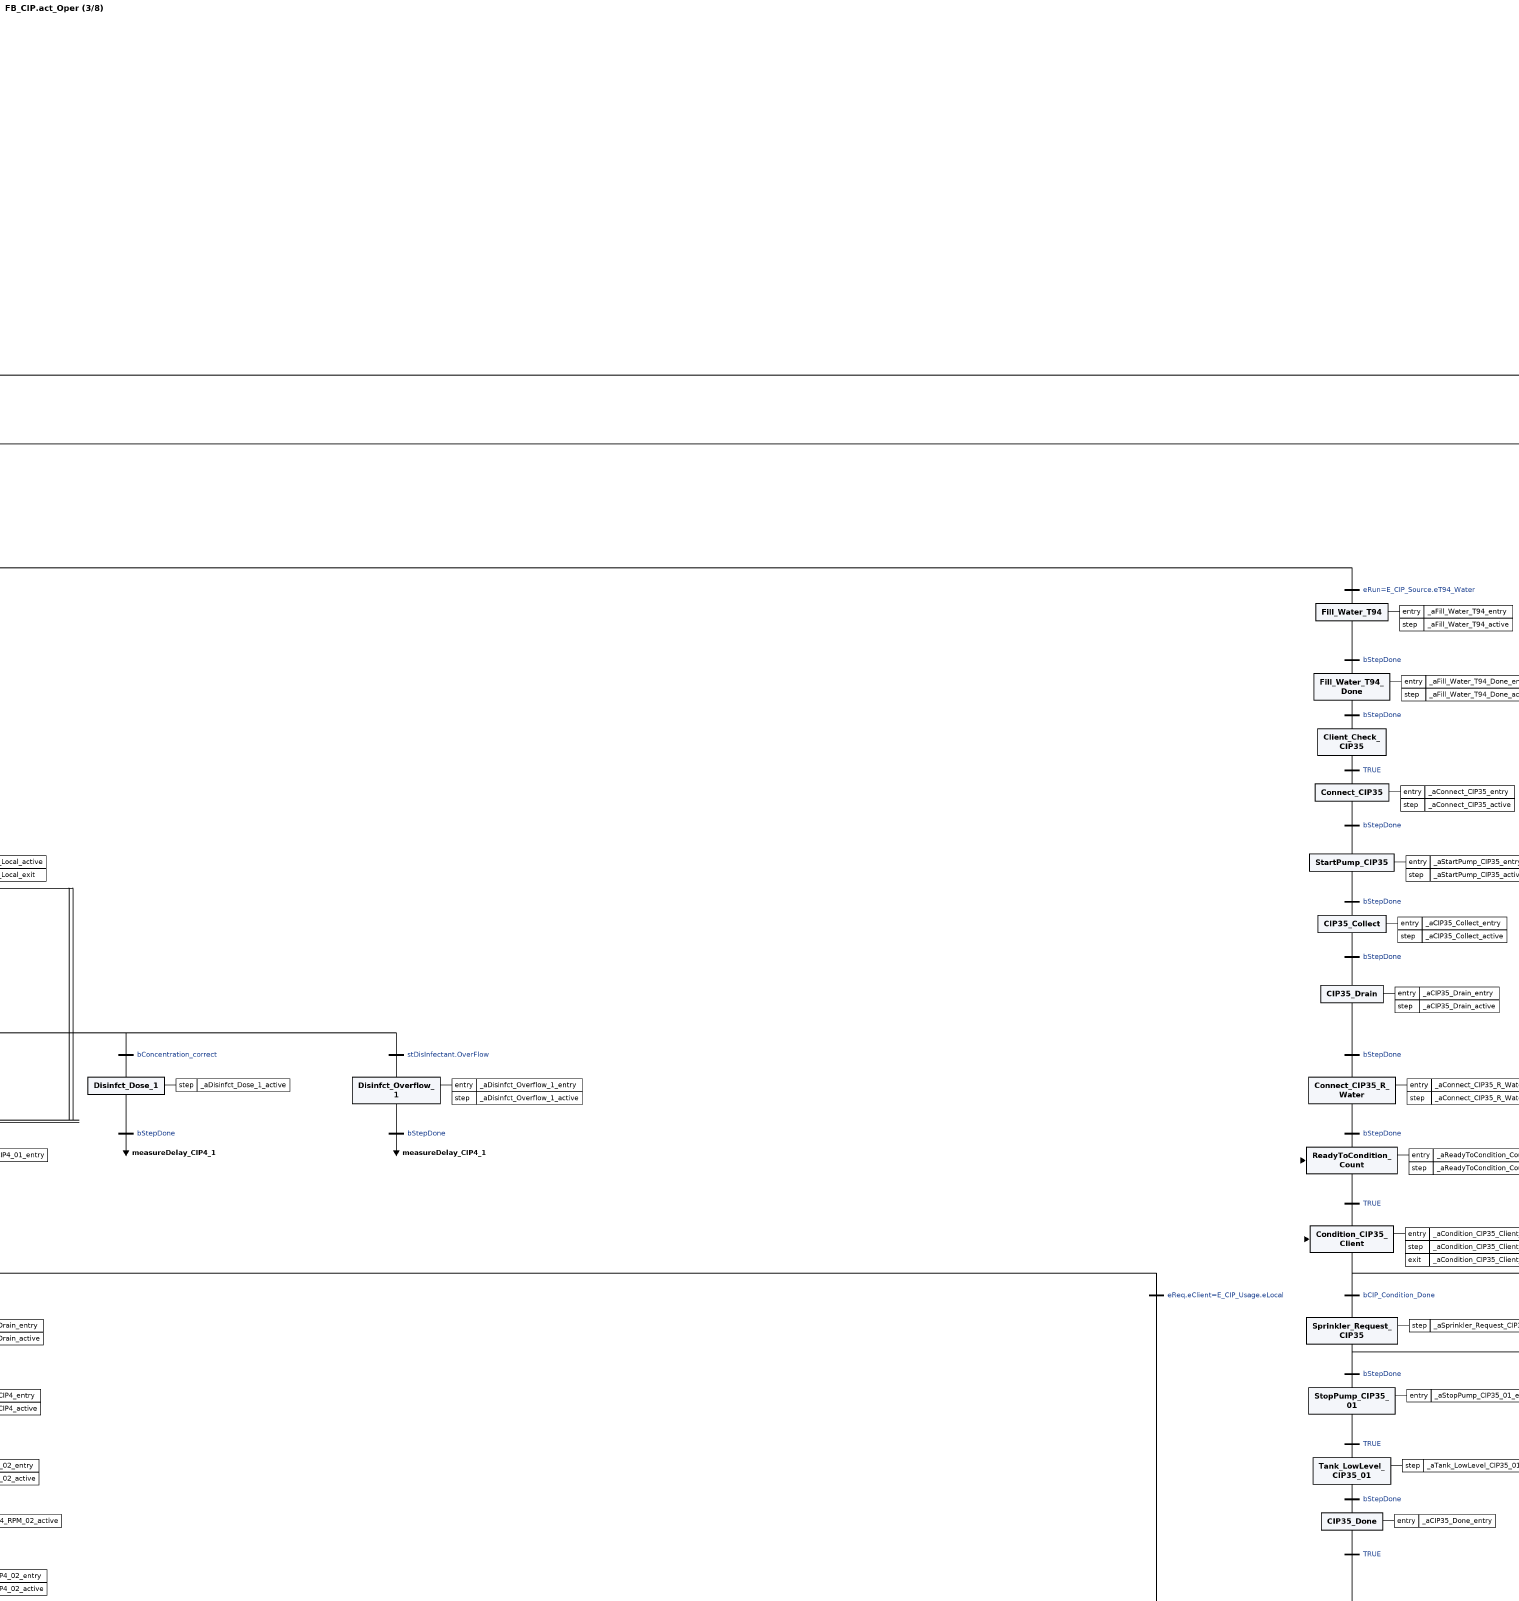
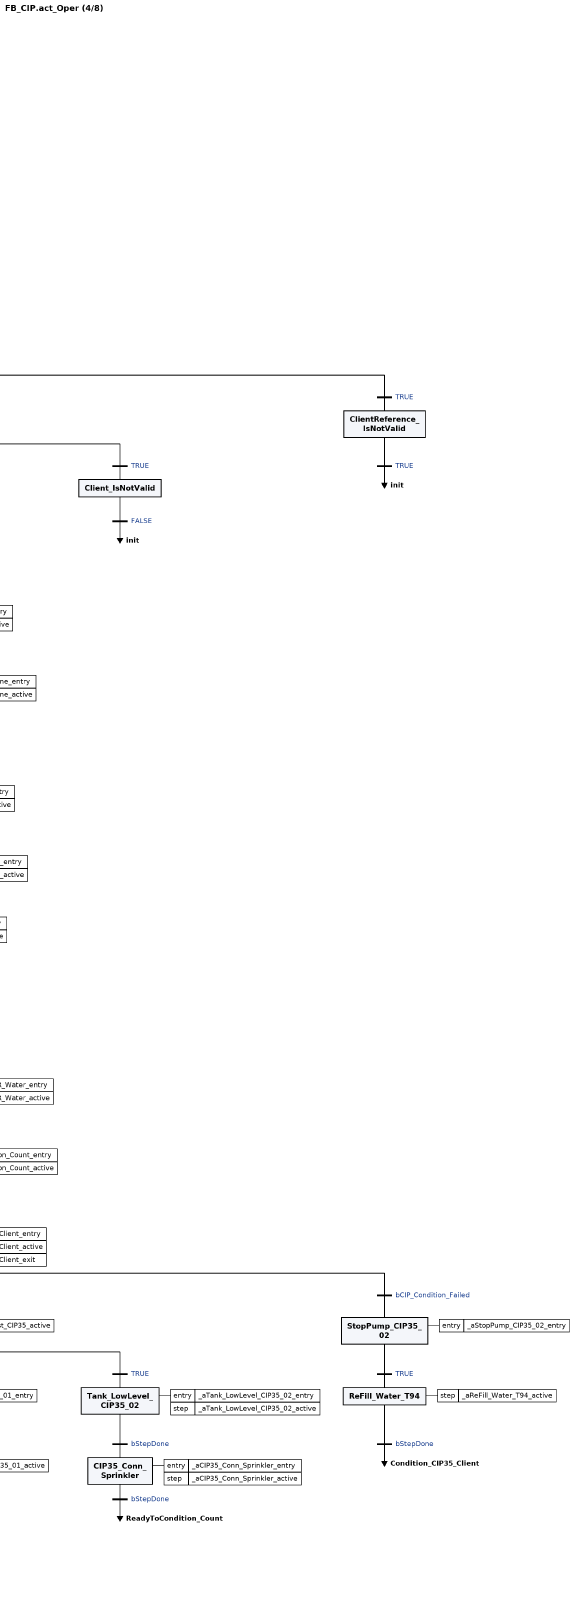
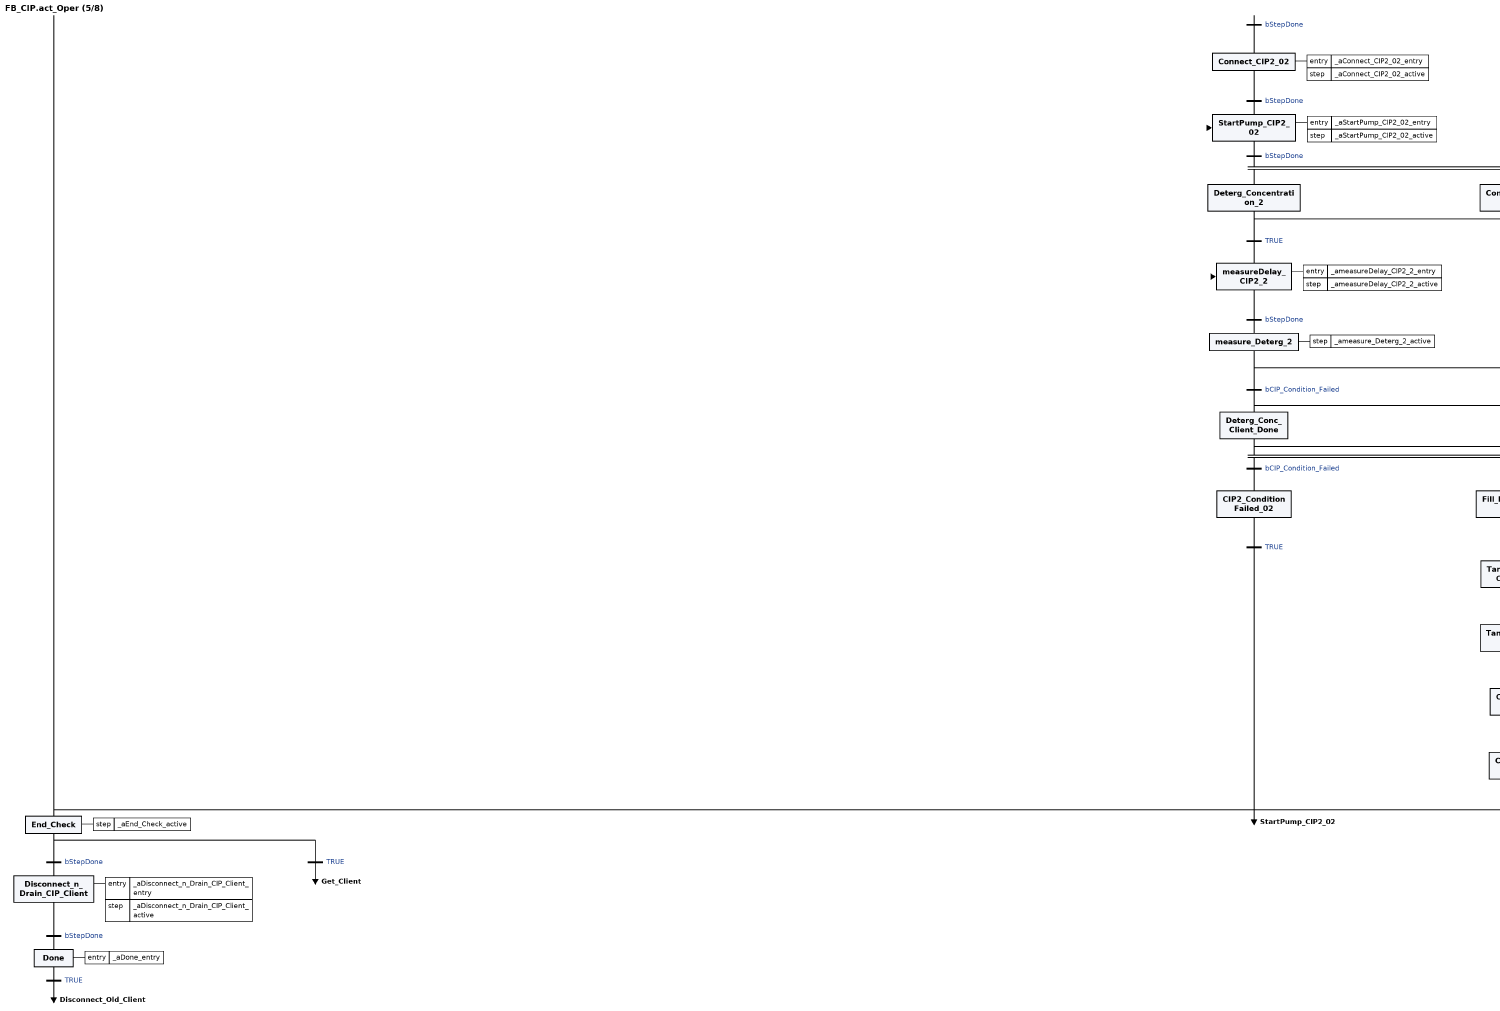
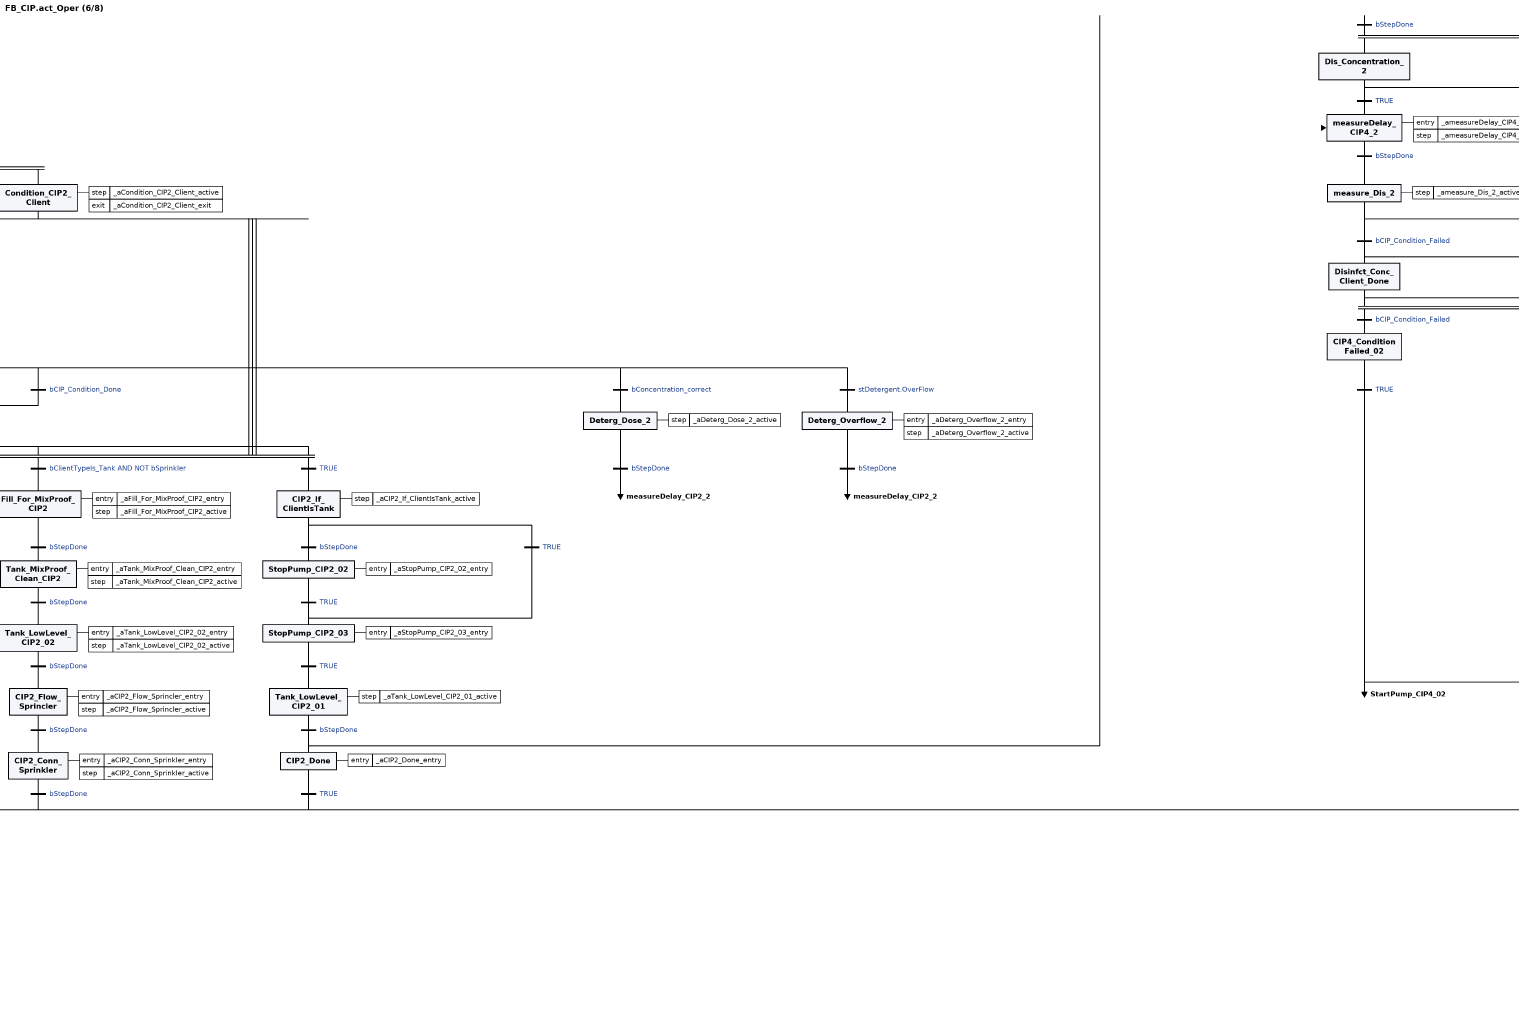
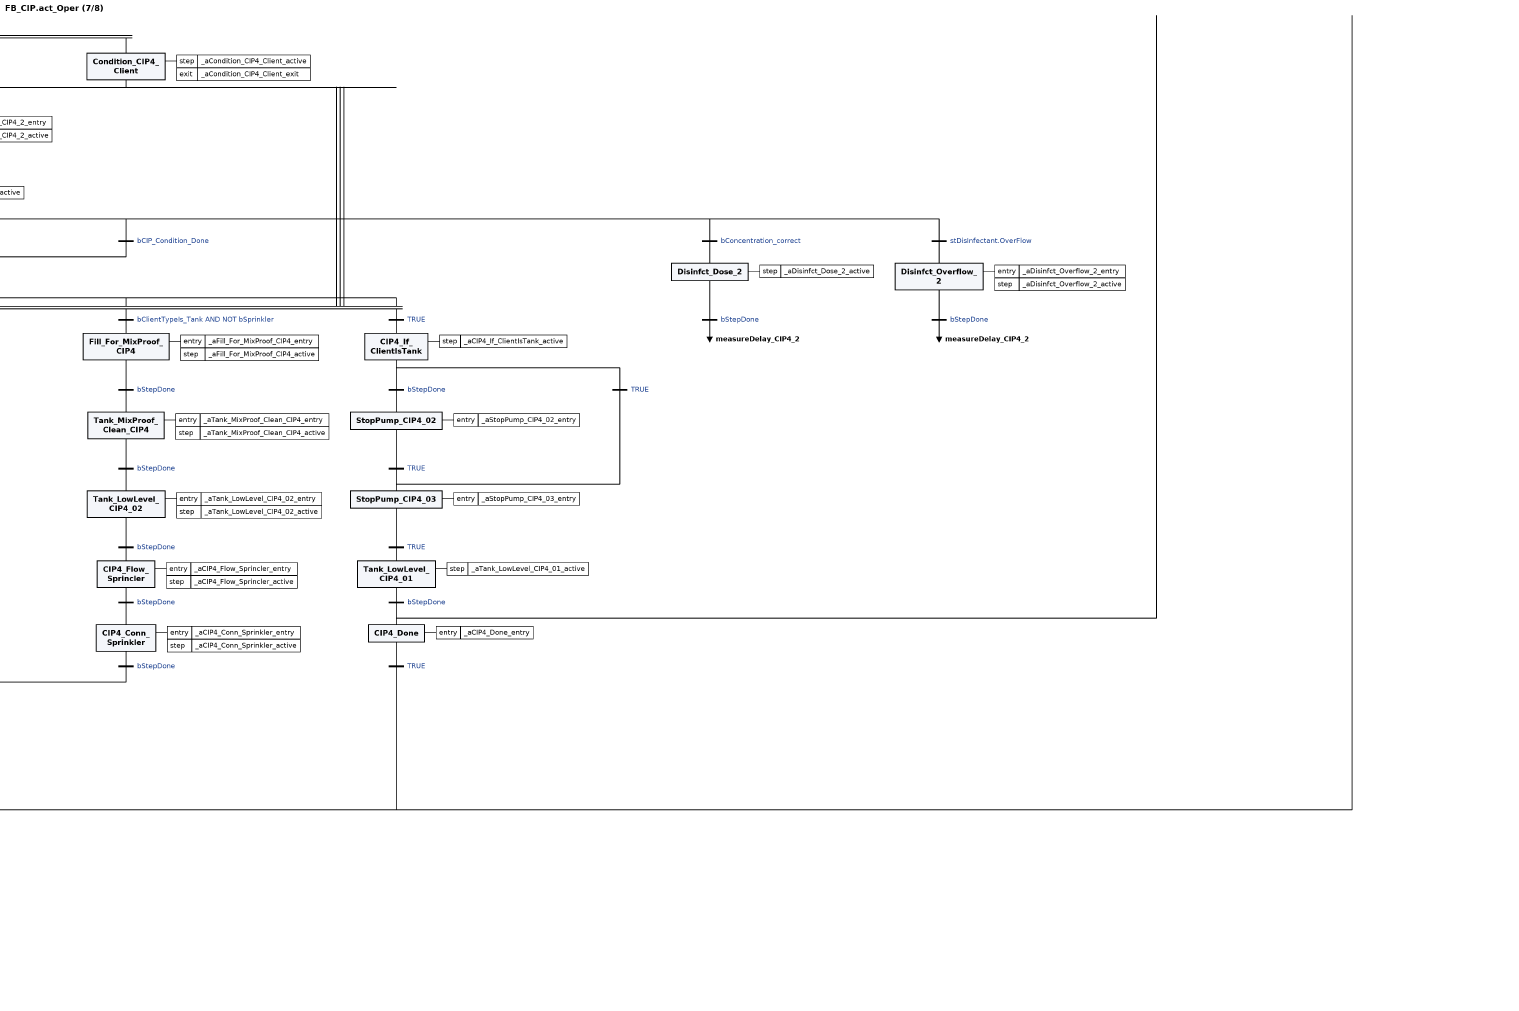
INITIAL_STEP init:
    _ainit_active(N);  // step action
    _ainit_exit(P0);  // exit action
END_STEP
TRANSITION FROM init TO Stop_Pump
    := TRUE;
END_TRANSITION
STEP Stop_Pump:
    _aStop_Pump_entry(P1);  // entry action
END_STEP
TRANSITION FROM Stop_Pump TO Set_Valves_ToDeafult
    := TRUE;
END_TRANSITION
STEP Set_Valves_ToDeafult:  // min time T#0.1s
    _aSet_Valves_ToDeafult_entry(P1);  // entry action
    _aSet_Valves_ToDeafult_active(N);  // step action
END_STEP
TRANSITION FROM Set_Valves_ToDeafult TO Waiting_Client_Drain_Done
    := bStepDone;
END_TRANSITION
STEP Waiting_Client_Drain_Done:  // min time T#0.1s
    _aWaiting_Client_Drain_Done_active(N);  // step action
END_STEP
TRANSITION FROM Waiting_Client_Drain_Done TO Disconnect_Old_Client
    := bStepDone;
END_TRANSITION
STEP Disconnect_Old_Client:
    _aDisconnect_Old_Client_entry(P1);  // entry action
END_STEP
TRANSITION FROM Disconnect_Old_Client TO Ready
    := TRUE;
END_TRANSITION
STEP Ready:
    _aReady_active(N);  // step action
    _aReady_exit(P0);  // exit action
END_STEP
TRANSITION FROM Ready TO Get_Client
    := bStepDone;
END_TRANSITION
STEP Get_Client:  // max time T#0.1s
    _aGet_Client_active(N);  // step action
    _aGet_Client_exit(P0);  // exit action
END_STEP
TRANSITION FROM Get_Client TO Client_Validation_check
    := bStepDone;
END_TRANSITION
TRANSITION FROM Get_Client TO ClientReference_IsNotValid
    := TRUE;
END_TRANSITION
STEP ClientReference_IsNotValid:  // min time T#2s
END_STEP
TRANSITION FROM ClientReference_IsNotValid TO init
    := TRUE;
END_TRANSITION
STEP Client_Validation_check:
    _aClient_Validation_check_active(N);  // step action
END_STEP
TRANSITION FROM Client_Validation_check TO TriBlender_Selection
    := bStepDone;
END_TRANSITION
STEP TriBlender_Selection:
    _aTriBlender_Selection_entry(P1);  // entry action
    _aTriBlender_Selection_active(N);  // step action
END_STEP
TRANSITION FROM TriBlender_Selection TO ClientReference_IsValid
    := bStepDone;
END_TRANSITION
TRANSITION FROM Client_Validation_check TO Client_IsNotValid
    := TRUE;
END_TRANSITION
STEP Client_IsNotValid:  // min time T#2s
END_STEP
TRANSITION FROM Client_IsNotValid TO init
    := FALSE;
END_TRANSITION
STEP ClientReference_IsValid:
    _aClientReference_IsValid_entry(P1);  // entry action
END_STEP
TRANSITION FROM ClientReference_IsValid TO Client_Check_01
    := eRun=E_CIP_Source.eT93_R_Water;
END_TRANSITION
// macro R_Water begins
STEP Client_Check_01:
END_STEP
TRANSITION FROM Client_Check_01 TO Fill_Water_T93
    := eReq.eClient<>E_CIP_Usage.eLocal;
END_TRANSITION
STEP Fill_Water_T93:
    _aFill_Water_T93_entry(P1);  // entry action
    _aFill_Water_T93_active(N);  // step action
END_STEP
TRANSITION FROM Fill_Water_T93 TO Fill_Water_T93_Done
    := bStepDone;
END_TRANSITION
STEP Fill_Water_T93_Done:
    _aFill_Water_T93_Done_entry(P1);  // entry action
    _aFill_Water_T93_Done_active(N);  // step action
END_STEP
TRANSITION FROM Fill_Water_T93_Done TO Client_tank_IsEmpty
    := bStepDone;
END_TRANSITION
STEP Client_tank_IsEmpty:  // min time T#5s
    _aClient_tank_IsEmpty_active(N);  // step action
END_STEP
TRANSITION FROM Client_tank_IsEmpty TO Connect_CIP1_Drain
    := bStepDone;
END_TRANSITION
STEP Connect_CIP1_Drain:
    _aConnect_CIP1_Drain_entry(P1);  // entry action
    _aConnect_CIP1_Drain_active(N);  // step action
END_STEP
TRANSITION FROM Connect_CIP1_Drain TO StartPump_CIP1_01
    := bStepDone;
END_TRANSITION
STEP StartPump_CIP1_01:
    _aStartPump_CIP1_01_entry(P1);  // entry action
    _aStartPump_CIP1_01_active(N);  // step action
END_STEP
TRANSITION FROM StartPump_CIP1_01 TO Condition_CIP1_Client
    := bStepDone;
END_TRANSITION
STEP Condition_CIP1_Client:
    _aCondition_CIP1_Client_entry(P1);  // entry action
    _aCondition_CIP1_Client_active(N);  // step action
    _aCondition_CIP1_Client_exit(P0);  // exit action
END_STEP
TRANSITION FROM Condition_CIP1_Client TO Sprinkler_Request_CIP1
    := bCIP_Condition_Done;
END_TRANSITION
STEP Sprinkler_Request_CIP1:
    _aSprinkler_Request_CIP1_active(N);  // step action
END_STEP
TRANSITION FROM Sprinkler_Request_CIP1 TO StopPump_CIP1_01
    := bStepDone;
END_TRANSITION
STEP StopPump_CIP1_01:
    _aStopPump_CIP1_01_entry(P1);  // entry action
END_STEP
TRANSITION FROM StopPump_CIP1_01 TO Tank_LowLevel_CIP1_01
    := TRUE;
END_TRANSITION
STEP Tank_LowLevel_CIP1_01:
    _aTank_LowLevel_CIP1_01_active(N);  // step action
END_STEP
TRANSITION FROM Tank_LowLevel_CIP1_01 TO CIP1_Done
    := bStepDone;
END_TRANSITION
TRANSITION FROM Sprinkler_Request_CIP1 TO Tank_LowLevel_CIP1_02
    := TRUE;
END_TRANSITION
STEP Tank_LowLevel_CIP1_02:
    _aTank_LowLevel_CIP1_02_entry(P1);  // entry action
    _aTank_LowLevel_CIP1_02_active(N);  // step action
END_STEP
TRANSITION FROM Tank_LowLevel_CIP1_02 TO CIP1_Conn_Sprinkler
    := bStepDone;
END_TRANSITION
STEP CIP1_Conn_Sprinkler:
    _aCIP1_Conn_Sprinkler_entry(P1);  // entry action
    _aCIP1_Conn_Sprinkler_active(N);  // step action
END_STEP
TRANSITION FROM CIP1_Conn_Sprinkler TO StartPump_CIP1_01
    := bStepDone;
END_TRANSITION
TRANSITION FROM Condition_CIP1_Client TO StopPump_CIP1_02
    := bCIP_Condition_Failed;
END_TRANSITION
STEP StopPump_CIP1_02:
    _aStopPump_CIP1_02_entry(P1);  // entry action
END_STEP
TRANSITION FROM StopPump_CIP1_02 TO ReFill_Water_T93
    := TRUE;
END_TRANSITION
STEP ReFill_Water_T93:
    _aReFill_Water_T93_active(N);  // step action
END_STEP
TRANSITION FROM ReFill_Water_T93 TO Condition_CIP1_Client
    := bStepDone;
END_TRANSITION
TRANSITION FROM Client_Check_01 TO CIP1_Done
    := eReq.eClient=E_CIP_Usage.eLocal;
END_TRANSITION
STEP CIP1_Done:  // min time T#2s
    _aCIP1_Done_entry(P1);  // entry action
END_STEP
TRANSITION FROM CIP1_Done TO End_Check
    := TRUE;
END_TRANSITION
TRANSITION FROM ClientReference_IsValid TO Fill_Water_T92
    := eRun=E_CIP_Source.eT92_Detergent;
END_TRANSITION
// macro Detergent begins
STEP Fill_Water_T92:
    _aFill_Water_T92_entry(P1);  // entry action
    _aFill_Water_T92_active(N);  // step action
END_STEP
TRANSITION FROM Fill_Water_T92 TO Connect_CIP2_01
    := bStepDone;
END_TRANSITION
STEP Connect_CIP2_01:
    _aConnect_CIP2_01_entry(P1);  // entry action
    _aConnect_CIP2_01_active(N);  // step action
END_STEP
TRANSITION FROM Connect_CIP2_01 TO Reset_Cond_Tm_CIP2_01
    := bStepDone;
END_TRANSITION
STEP Reset_Cond_Tm_CIP2_01:
    _aReset_Cond_Tm_CIP2_01_active(N);  // step action
END_STEP
TRANSITION FROM Reset_Cond_Tm_CIP2_01 TO CheckIf_CIP_Pump_Ready
    := TRUE;
END_TRANSITION
STEP CheckIf_CIP_Pump_Ready:
END_STEP
TRANSITION FROM CheckIf_CIP_Pump_Ready TO StartPump_CIP2_RPM_01
    := fb_PumpCIP.DriveReady;
END_TRANSITION
STEP StartPump_CIP2_RPM_01:
    _aStartPump_CIP2_RPM_01_active(N);  // step action
END_STEP
TRANSITION FROM StartPump_CIP2_RPM_01 TO StartPump_CIP2_01
    := bStepDone;
END_TRANSITION
STEP StartPump_CIP2_01:  // min time T#2s
    _aStartPump_CIP2_01_entry(P1);  // entry action
    _aStartPump_CIP2_01_active(N);  // step action
END_STEP
TRANSITION FROM StartPump_CIP2_01 TO (Deterg_Concentration_1, Condition_CIP2_Local)
    := bStepDone;
END_TRANSITION
STEP Deterg_Concentration_1:
END_STEP
TRANSITION FROM Deterg_Concentration_1 TO measureDelay_CIP2_1
    := TRUE;
END_TRANSITION
STEP measureDelay_CIP2_1:
    _ameasureDelay_CIP2_1_entry(P1);  // entry action
    _ameasureDelay_CIP2_1_active(N);  // step action
END_STEP
TRANSITION FROM measureDelay_CIP2_1 TO measure_Deterg
    := bStepDone;
END_TRANSITION
STEP measure_Deterg:  // min time t#1s
    _ameasure_Deterg_active(N);  // step action
END_STEP
TRANSITION FROM measure_Deterg TO Deterg_Conc_Local_Done
    := bCIP_Condition_Failed;
END_TRANSITION
TRANSITION FROM measure_Deterg TO Deterg_Conc_Local_Done
    := bCIP_Condition_Done;
END_TRANSITION
TRANSITION FROM measure_Deterg TO Deterg_Dose_1
    := bConcentration_correct;
END_TRANSITION
STEP Deterg_Dose_1:
    _aDeterg_Dose_1_active(N);  // step action
END_STEP
TRANSITION FROM Deterg_Dose_1 TO measureDelay_CIP2_1
    := bStepDone;
END_TRANSITION
TRANSITION FROM measure_Deterg TO Deterg_Overflow_1
    := stDetergent.OverFlow;
END_TRANSITION
STEP Deterg_Overflow_1:
    _aDeterg_Overflow_1_entry(P1);  // entry action
    _aDeterg_Overflow_1_active(N);  // step action
END_STEP
TRANSITION FROM Deterg_Overflow_1 TO measureDelay_CIP2_1
    := bStepDone;
END_TRANSITION
STEP Deterg_Conc_Local_Done:
END_STEP
STEP Condition_CIP2_Local:
    _aCondition_CIP2_Local_active(N);  // step action
    _aCondition_CIP2_Local_exit(P0);  // exit action
END_STEP
TRANSITION FROM (Deterg_Conc_Local_Done, Condition_CIP2_Local) TO CIP2_ConditionFailed_01
    := bCIP_Condition_Failed;
END_TRANSITION
STEP CIP2_ConditionFailed_01:
END_STEP
TRANSITION FROM CIP2_ConditionFailed_01 TO StartPump_CIP2_01
    := TRUE;
END_TRANSITION
TRANSITION FROM (Deterg_Conc_Local_Done, Condition_CIP2_Local) TO StopPump_CIP2_01
    := bCIP_Condition_Done;
END_TRANSITION
STEP StopPump_CIP2_01:
    _aStopPump_CIP2_01_entry(P1);  // entry action
END_STEP
TRANSITION FROM StopPump_CIP2_01 TO Client_Check_CIP2
    := TRUE;
END_TRANSITION
STEP Client_Check_CIP2:
END_STEP
TRANSITION FROM Client_Check_CIP2 TO Connect_CIP2_Drain
    := eReq.eClient<>E_CIP_Usage.eLocal;
END_TRANSITION
STEP Connect_CIP2_Drain:
    _aConnect_CIP2_Drain_entry(P1);  // entry action
    _aConnect_CIP2_Drain_active(N);  // step action
END_STEP
TRANSITION FROM Connect_CIP2_Drain TO StartPump_CIP2_RPM_02
    := bStepDone;
END_TRANSITION
STEP StartPump_CIP2_RPM_02:
    _aStartPump_CIP2_RPM_02_entry(P1);  // entry action
    _aStartPump_CIP2_RPM_02_active(N);  // step action
END_STEP
TRANSITION FROM StartPump_CIP2_RPM_02 TO Fill_Solution_CIP2
    := bStepDone;
END_TRANSITION
STEP Fill_Solution_CIP2:
    _aFill_Solution_CIP2_active(N);  // step action
END_STEP
TRANSITION FROM Fill_Solution_CIP2 TO Connect_CIP2_02
    := bStepDone;
END_TRANSITION
STEP Connect_CIP2_02:
    _aConnect_CIP2_02_entry(P1);  // entry action
    _aConnect_CIP2_02_active(N);  // step action
END_STEP
TRANSITION FROM Connect_CIP2_02 TO StartPump_CIP2_02
    := bStepDone;
END_TRANSITION
STEP StartPump_CIP2_02:  // min time T#2s
    _aStartPump_CIP2_02_entry(P1);  // entry action
    _aStartPump_CIP2_02_active(N);  // step action
END_STEP
TRANSITION FROM StartPump_CIP2_02 TO (Deterg_Concentration_2, Condition_CIP2_Client)
    := bStepDone;
END_TRANSITION
STEP Deterg_Concentration_2:
END_STEP
TRANSITION FROM Deterg_Concentration_2 TO measureDelay_CIP2_2
    := TRUE;
END_TRANSITION
STEP measureDelay_CIP2_2:
    _ameasureDelay_CIP2_2_entry(P1);  // entry action
    _ameasureDelay_CIP2_2_active(N);  // step action
END_STEP
TRANSITION FROM measureDelay_CIP2_2 TO measure_Deterg_2
    := bStepDone;
END_TRANSITION
STEP measure_Deterg_2:  // min time t#1s
    _ameasure_Deterg_2_active(N);  // step action
END_STEP
TRANSITION FROM measure_Deterg_2 TO Deterg_Conc_Client_Done
    := bCIP_Condition_Failed;
END_TRANSITION
TRANSITION FROM measure_Deterg_2 TO Deterg_Conc_Client_Done
    := bCIP_Condition_Done;
END_TRANSITION
TRANSITION FROM measure_Deterg_2 TO Deterg_Dose_2
    := bConcentration_correct;
END_TRANSITION
STEP Deterg_Dose_2:
    _aDeterg_Dose_2_active(N);  // step action
END_STEP
TRANSITION FROM Deterg_Dose_2 TO measureDelay_CIP2_2
    := bStepDone;
END_TRANSITION
TRANSITION FROM measure_Deterg_2 TO Deterg_Overflow_2
    := stDetergent.OverFlow;
END_TRANSITION
STEP Deterg_Overflow_2:
    _aDeterg_Overflow_2_entry(P1);  // entry action
    _aDeterg_Overflow_2_active(N);  // step action
END_STEP
TRANSITION FROM Deterg_Overflow_2 TO measureDelay_CIP2_2
    := bStepDone;
END_TRANSITION
STEP Deterg_Conc_Client_Done:
END_STEP
STEP Condition_CIP2_Client:
    _aCondition_CIP2_Client_active(N);  // step action
    _aCondition_CIP2_Client_exit(P0);  // exit action
END_STEP
TRANSITION FROM (Deterg_Conc_Client_Done, Condition_CIP2_Client) TO CIP2_ConditionFailed_02
    := bCIP_Condition_Failed;
END_TRANSITION
STEP CIP2_ConditionFailed_02:
END_STEP
TRANSITION FROM CIP2_ConditionFailed_02 TO StartPump_CIP2_02
    := TRUE;
END_TRANSITION
TRANSITION FROM (Deterg_Conc_Client_Done, Condition_CIP2_Client) TO Fill_For_MixProof_CIP2
    := bClientTypeIs_Tank AND NOT bSprinkler;
END_TRANSITION
STEP Fill_For_MixProof_CIP2:
    _aFill_For_MixProof_CIP2_entry(P1);  // entry action
    _aFill_For_MixProof_CIP2_active(N);  // step action
END_STEP
TRANSITION FROM Fill_For_MixProof_CIP2 TO Tank_MixProof_Clean_CIP2
    := bStepDone;
END_TRANSITION
STEP Tank_MixProof_Clean_CIP2:
    _aTank_MixProof_Clean_CIP2_entry(P1);  // entry action
    _aTank_MixProof_Clean_CIP2_active(N);  // step action
END_STEP
TRANSITION FROM Tank_MixProof_Clean_CIP2 TO Tank_LowLevel_CIP2_02
    := bStepDone;
END_TRANSITION
STEP Tank_LowLevel_CIP2_02:
    _aTank_LowLevel_CIP2_02_entry(P1);  // entry action
    _aTank_LowLevel_CIP2_02_active(N);  // step action
END_STEP
TRANSITION FROM Tank_LowLevel_CIP2_02 TO CIP2_Flow_Sprincler
    := bStepDone;
END_TRANSITION
STEP CIP2_Flow_Sprincler:
    _aCIP2_Flow_Sprincler_entry(P1);  // entry action
    _aCIP2_Flow_Sprincler_active(N);  // step action
END_STEP
TRANSITION FROM CIP2_Flow_Sprincler TO CIP2_Conn_Sprinkler
    := bStepDone;
END_TRANSITION
STEP CIP2_Conn_Sprinkler:
    _aCIP2_Conn_Sprinkler_entry(P1);  // entry action
    _aCIP2_Conn_Sprinkler_active(N);  // step action
END_STEP
TRANSITION FROM CIP2_Conn_Sprinkler TO StartPump_CIP2_02
    := bStepDone;
END_TRANSITION
TRANSITION FROM (Deterg_Conc_Client_Done, Condition_CIP2_Client) TO CIP2_If_ClientIsTank
    := TRUE;
END_TRANSITION
STEP CIP2_If_ClientIsTank:
    _aCIP2_If_ClientIsTank_active(N);  // step action
END_STEP
TRANSITION FROM CIP2_If_ClientIsTank TO StopPump_CIP2_02
    := bStepDone;
END_TRANSITION
STEP StopPump_CIP2_02:
    _aStopPump_CIP2_02_entry(P1);  // entry action
END_STEP
TRANSITION FROM StopPump_CIP2_02 TO StopPump_CIP2_03
    := TRUE;
END_TRANSITION
TRANSITION FROM CIP2_If_ClientIsTank TO StopPump_CIP2_03
    := TRUE;
END_TRANSITION
STEP StopPump_CIP2_03:
    _aStopPump_CIP2_03_entry(P1);  // entry action
END_STEP
TRANSITION FROM StopPump_CIP2_03 TO Tank_LowLevel_CIP2_01
    := TRUE;
END_TRANSITION
STEP Tank_LowLevel_CIP2_01:
    _aTank_LowLevel_CIP2_01_active(N);  // step action
END_STEP
TRANSITION FROM Tank_LowLevel_CIP2_01 TO CIP2_Done
    := bStepDone;
END_TRANSITION
TRANSITION FROM Client_Check_CIP2 TO CIP2_Done
    := eReq.eClient=E_CIP_Usage.eLocal;
END_TRANSITION
STEP CIP2_Done:  // min time T#2s
    _aCIP2_Done_entry(P1);  // entry action
END_STEP
TRANSITION FROM CIP2_Done TO End_Check
    := TRUE;
END_TRANSITION
TRANSITION FROM ClientReference_IsValid TO Fill_Water_T91
    := eRun=E_CIP_Source.eT91_Sanitation;
END_TRANSITION
// macro DisInfection begins
STEP Fill_Water_T91:
    _aFill_Water_T91_entry(P1);  // entry action
    _aFill_Water_T91_active(N);  // step action
END_STEP
TRANSITION FROM Fill_Water_T91 TO Connect_CIP4_01
    := bStepDone;
END_TRANSITION
STEP Connect_CIP4_01:
    _aConnect_CIP4_01_entry(P1);  // entry action
    _aConnect_CIP4_01_active(N);  // step action
END_STEP
TRANSITION FROM Connect_CIP4_01 TO StartPump_CIP4_RPM_01
    := bStepDone;
END_TRANSITION
STEP StartPump_CIP4_RPM_01:
    _aStartPump_CIP4_RPM_01_active(N);  // step action
END_STEP
TRANSITION FROM StartPump_CIP4_RPM_01 TO StartPump_CIP4_01
    := bStepDone;
END_TRANSITION
STEP StartPump_CIP4_01:  // min time T#3s
    _aStartPump_CIP4_01_entry(P1);  // entry action
    _aStartPump_CIP4_01_active(N);  // step action
END_STEP
TRANSITION FROM StartPump_CIP4_01 TO (Dis_Concentration_1, Condition_CIP4_Local)
    := bStepDone;
END_TRANSITION
STEP Dis_Concentration_1:
END_STEP
TRANSITION FROM Dis_Concentration_1 TO measureDelay_CIP4_1
    := TRUE;
END_TRANSITION
STEP measureDelay_CIP4_1:
    _ameasureDelay_CIP4_1_entry(P1);  // entry action
    _ameasureDelay_CIP4_1_active(N);  // step action
END_STEP
TRANSITION FROM measureDelay_CIP4_1 TO measure_Dis
    := bStepDone;
END_TRANSITION
STEP measure_Dis:  // min time t#1s
    _ameasure_Dis_active(N);  // step action
END_STEP
TRANSITION FROM measure_Dis TO Disinfct_Conc_Local_Done
    := bCIP_Condition_Failed;
END_TRANSITION
TRANSITION FROM measure_Dis TO Disinfct_Conc_Local_Done
    := bCIP_Condition_Done;
END_TRANSITION
TRANSITION FROM measure_Dis TO Disinfct_Dose_1
    := bConcentration_correct;
END_TRANSITION
STEP Disinfct_Dose_1:
    _aDisinfct_Dose_1_active(N);  // step action
END_STEP
TRANSITION FROM Disinfct_Dose_1 TO measureDelay_CIP4_1
    := bStepDone;
END_TRANSITION
TRANSITION FROM measure_Dis TO Disinfct_Overflow_1
    := stDisInfectant.OverFlow;
END_TRANSITION
STEP Disinfct_Overflow_1:
    _aDisinfct_Overflow_1_entry(P1);  // entry action
    _aDisinfct_Overflow_1_active(N);  // step action
END_STEP
TRANSITION FROM Disinfct_Overflow_1 TO measureDelay_CIP4_1
    := bStepDone;
END_TRANSITION
STEP Disinfct_Conc_Local_Done:
END_STEP
STEP Condition_CIP4_Local:
    _aCondition_CIP4_Local_active(N);  // step action
    _aCondition_CIP4_Local_exit(P0);  // exit action
END_STEP
TRANSITION FROM (Disinfct_Conc_Local_Done, Condition_CIP4_Local) TO CIP4_ConditionFailed_01
    := bCIP_Condition_Failed;
END_TRANSITION
STEP CIP4_ConditionFailed_01:
END_STEP
TRANSITION FROM CIP4_ConditionFailed_01 TO StartPump_CIP4_01
    := TRUE;
END_TRANSITION
TRANSITION FROM (Disinfct_Conc_Local_Done, Condition_CIP4_Local) TO StopPump_CIP4_01
    := bCIP_Condition_Done;
END_TRANSITION
STEP StopPump_CIP4_01:  // min time T#5s
    _aStopPump_CIP4_01_entry(P1);  // entry action
END_STEP
TRANSITION FROM StopPump_CIP4_01 TO Client_Check_CIP4
    := TRUE;
END_TRANSITION
STEP Client_Check_CIP4:
END_STEP
TRANSITION FROM Client_Check_CIP4 TO Connect_CIP4_Drain
    := eReq.eClient<>E_CIP_Usage.eLocal;
END_TRANSITION
STEP Connect_CIP4_Drain:
    _aConnect_CIP4_Drain_entry(P1);  // entry action
    _aConnect_CIP4_Drain_active(N);  // step action
END_STEP
TRANSITION FROM Connect_CIP4_Drain TO Fill_Solution_CIP4
    := bStepDone;
END_TRANSITION
STEP Fill_Solution_CIP4:
    _aFill_Solution_CIP4_entry(P1);  // entry action
    _aFill_Solution_CIP4_active(N);  // step action
END_STEP
TRANSITION FROM Fill_Solution_CIP4 TO Connect_CIP4_02
    := bStepDone;
END_TRANSITION
STEP Connect_CIP4_02:
    _aConnect_CIP4_02_entry(P1);  // entry action
    _aConnect_CIP4_02_active(N);  // step action
END_STEP
TRANSITION FROM Connect_CIP4_02 TO StartPump_CIP4_RPM_02
    := bStepDone;
END_TRANSITION
STEP StartPump_CIP4_RPM_02:
    _aStartPump_CIP4_RPM_02_active(N);  // step action
END_STEP
TRANSITION FROM StartPump_CIP4_RPM_02 TO StartPump_CIP4_02
    := bStepDone;
END_TRANSITION
STEP StartPump_CIP4_02:  // min time T#1s
    _aStartPump_CIP4_02_entry(P1);  // entry action
    _aStartPump_CIP4_02_active(N);  // step action
END_STEP
TRANSITION FROM StartPump_CIP4_02 TO (Dis_Concentration_2, Condition_CIP4_Client)
    := bStepDone;
END_TRANSITION
STEP Dis_Concentration_2:
END_STEP
TRANSITION FROM Dis_Concentration_2 TO measureDelay_CIP4_2
    := TRUE;
END_TRANSITION
STEP measureDelay_CIP4_2:
    _ameasureDelay_CIP4_2_entry(P1);  // entry action
    _ameasureDelay_CIP4_2_active(N);  // step action
END_STEP
TRANSITION FROM measureDelay_CIP4_2 TO measure_Dis_2
    := bStepDone;
END_TRANSITION
STEP measure_Dis_2:  // min time t#1s
    _ameasure_Dis_2_active(N);  // step action
END_STEP
TRANSITION FROM measure_Dis_2 TO Disinfct_Conc_Client_Done
    := bCIP_Condition_Failed;
END_TRANSITION
TRANSITION FROM measure_Dis_2 TO Disinfct_Conc_Client_Done
    := bCIP_Condition_Done;
END_TRANSITION
TRANSITION FROM measure_Dis_2 TO Disinfct_Dose_2
    := bConcentration_correct;
END_TRANSITION
STEP Disinfct_Dose_2:
    _aDisinfct_Dose_2_active(N);  // step action
END_STEP
TRANSITION FROM Disinfct_Dose_2 TO measureDelay_CIP4_2
    := bStepDone;
END_TRANSITION
TRANSITION FROM measure_Dis_2 TO Disinfct_Overflow_2
    := stDisInfectant.OverFlow;
END_TRANSITION
STEP Disinfct_Overflow_2:
    _aDisinfct_Overflow_2_entry(P1);  // entry action
    _aDisinfct_Overflow_2_active(N);  // step action
END_STEP
TRANSITION FROM Disinfct_Overflow_2 TO measureDelay_CIP4_2
    := bStepDone;
END_TRANSITION
STEP Disinfct_Conc_Client_Done:
END_STEP
STEP Condition_CIP4_Client:
    _aCondition_CIP4_Client_active(N);  // step action
    _aCondition_CIP4_Client_exit(P0);  // exit action
END_STEP
TRANSITION FROM (Disinfct_Conc_Client_Done, Condition_CIP4_Client) TO CIP4_ConditionFailed_02
    := bCIP_Condition_Failed;
END_TRANSITION
STEP CIP4_ConditionFailed_02:
END_STEP
TRANSITION FROM CIP4_ConditionFailed_02 TO StartPump_CIP4_02
    := TRUE;
END_TRANSITION
TRANSITION FROM (Disinfct_Conc_Client_Done, Condition_CIP4_Client) TO Fill_For_MixProof_CIP4
    := bClientTypeIs_Tank AND NOT bSprinkler;
END_TRANSITION
STEP Fill_For_MixProof_CIP4:
    _aFill_For_MixProof_CIP4_entry(P1);  // entry action
    _aFill_For_MixProof_CIP4_active(N);  // step action
END_STEP
TRANSITION FROM Fill_For_MixProof_CIP4 TO Tank_MixProof_Clean_CIP4
    := bStepDone;
END_TRANSITION
STEP Tank_MixProof_Clean_CIP4:
    _aTank_MixProof_Clean_CIP4_entry(P1);  // entry action
    _aTank_MixProof_Clean_CIP4_active(N);  // step action
END_STEP
TRANSITION FROM Tank_MixProof_Clean_CIP4 TO Tank_LowLevel_CIP4_02
    := bStepDone;
END_TRANSITION
STEP Tank_LowLevel_CIP4_02:
    _aTank_LowLevel_CIP4_02_entry(P1);  // entry action
    _aTank_LowLevel_CIP4_02_active(N);  // step action
END_STEP
TRANSITION FROM Tank_LowLevel_CIP4_02 TO CIP4_Flow_Sprincler
    := bStepDone;
END_TRANSITION
STEP CIP4_Flow_Sprincler:
    _aCIP4_Flow_Sprincler_entry(P1);  // entry action
    _aCIP4_Flow_Sprincler_active(N);  // step action
END_STEP
TRANSITION FROM CIP4_Flow_Sprincler TO CIP4_Conn_Sprinkler
    := bStepDone;
END_TRANSITION
STEP CIP4_Conn_Sprinkler:
    _aCIP4_Conn_Sprinkler_entry(P1);  // entry action
    _aCIP4_Conn_Sprinkler_active(N);  // step action
END_STEP
TRANSITION FROM CIP4_Conn_Sprinkler TO StartPump_CIP4_02
    := bStepDone;
END_TRANSITION
TRANSITION FROM (Disinfct_Conc_Client_Done, Condition_CIP4_Client) TO CIP4_If_ClientIsTank
    := TRUE;
END_TRANSITION
STEP CIP4_If_ClientIsTank:
    _aCIP4_If_ClientIsTank_active(N);  // step action
END_STEP
TRANSITION FROM CIP4_If_ClientIsTank TO StopPump_CIP4_02
    := bStepDone;
END_TRANSITION
STEP StopPump_CIP4_02:  // min time T#2s
    _aStopPump_CIP4_02_entry(P1);  // entry action
END_STEP
TRANSITION FROM StopPump_CIP4_02 TO StopPump_CIP4_03
    := TRUE;
END_TRANSITION
TRANSITION FROM CIP4_If_ClientIsTank TO StopPump_CIP4_03
    := TRUE;
END_TRANSITION
STEP StopPump_CIP4_03:
    _aStopPump_CIP4_03_entry(P1);  // entry action
END_STEP
TRANSITION FROM StopPump_CIP4_03 TO Tank_LowLevel_CIP4_01
    := TRUE;
END_TRANSITION
STEP Tank_LowLevel_CIP4_01:
    _aTank_LowLevel_CIP4_01_active(N);  // step action
END_STEP
TRANSITION FROM Tank_LowLevel_CIP4_01 TO CIP4_Done
    := bStepDone;
END_TRANSITION
TRANSITION FROM Client_Check_CIP4 TO CIP4_Done
    := eReq.eClient=E_CIP_Usage.eLocal;
END_TRANSITION
STEP CIP4_Done:  // min time T#2s
    _aCIP4_Done_entry(P1);  // entry action
END_STEP
TRANSITION FROM CIP4_Done TO End_Check
    := TRUE;
END_TRANSITION
TRANSITION FROM ClientReference_IsValid TO Fill_Water_T94
    := eRun=E_CIP_Source.eT94_Water;
END_TRANSITION
// macro Water begins
STEP Fill_Water_T94:
    _aFill_Water_T94_entry(P1);  // entry action
    _aFill_Water_T94_active(N);  // step action
END_STEP
TRANSITION FROM Fill_Water_T94 TO Fill_Water_T94_Done
    := bStepDone;
END_TRANSITION
STEP Fill_Water_T94_Done:
    _aFill_Water_T94_Done_entry(P1);  // entry action
    _aFill_Water_T94_Done_active(N);  // step action
END_STEP
TRANSITION FROM Fill_Water_T94_Done TO Client_Check_CIP35
    := bStepDone;
END_TRANSITION
STEP Client_Check_CIP35:
END_STEP
TRANSITION FROM Client_Check_CIP35 TO Connect_CIP35
    := TRUE;
END_TRANSITION
STEP Connect_CIP35:
    _aConnect_CIP35_entry(P1);  // entry action
    _aConnect_CIP35_active(N);  // step action
END_STEP
TRANSITION FROM Connect_CIP35 TO StartPump_CIP35
    := bStepDone;
END_TRANSITION
STEP StartPump_CIP35:  // min time T#3s
    _aStartPump_CIP35_entry(P1);  // entry action
    _aStartPump_CIP35_active(N);  // step action
END_STEP
TRANSITION FROM StartPump_CIP35 TO CIP35_Collect
    := bStepDone;
END_TRANSITION
STEP CIP35_Collect:  // min time T#5s
    _aCIP35_Collect_entry(P1);  // entry action
    _aCIP35_Collect_active(N);  // step action
END_STEP
TRANSITION FROM CIP35_Collect TO CIP35_Drain
    := bStepDone;
END_TRANSITION
STEP CIP35_Drain:  // min time T#5s
    _aCIP35_Drain_entry(P1);  // entry action
    _aCIP35_Drain_active(N);  // step action
END_STEP
TRANSITION FROM CIP35_Drain TO Connect_CIP35_R_Water
    := bStepDone;
END_TRANSITION
STEP Connect_CIP35_R_Water:  // min time T#5s
    _aConnect_CIP35_R_Water_entry(P1);  // entry action
    _aConnect_CIP35_R_Water_active(N);  // step action
END_STEP
TRANSITION FROM Connect_CIP35_R_Water TO ReadyToCondition_Count
    := bStepDone;
END_TRANSITION
STEP ReadyToCondition_Count:
    _aReadyToCondition_Count_entry(P1);  // entry action
    _aReadyToCondition_Count_active(N);  // step action
END_STEP
TRANSITION FROM ReadyToCondition_Count TO Condition_CIP35_Client
    := TRUE;
END_TRANSITION
STEP Condition_CIP35_Client:
    _aCondition_CIP35_Client_entry(P1);  // entry action
    _aCondition_CIP35_Client_active(N);  // step action
    _aCondition_CIP35_Client_exit(P0);  // exit action
END_STEP
TRANSITION FROM Condition_CIP35_Client TO Sprinkler_Request_CIP35
    := bCIP_Condition_Done;
END_TRANSITION
STEP Sprinkler_Request_CIP35:
    _aSprinkler_Request_CIP35_active(N);  // step action
END_STEP
TRANSITION FROM Sprinkler_Request_CIP35 TO StopPump_CIP35_01
    := bStepDone;
END_TRANSITION
STEP StopPump_CIP35_01:
    _aStopPump_CIP35_01_entry(P1);  // entry action
END_STEP
TRANSITION FROM StopPump_CIP35_01 TO Tank_LowLevel_CIP35_01
    := TRUE;
END_TRANSITION
TRANSITION FROM Sprinkler_Request_CIP35 TO Tank_LowLevel_CIP35_02
    := TRUE;
END_TRANSITION
STEP Tank_LowLevel_CIP35_02:
    _aTank_LowLevel_CIP35_02_entry(P1);  // entry action
    _aTank_LowLevel_CIP35_02_active(N);  // step action
END_STEP
TRANSITION FROM Tank_LowLevel_CIP35_02 TO CIP35_Conn_Sprinkler
    := bStepDone;
END_TRANSITION
STEP CIP35_Conn_Sprinkler:
    _aCIP35_Conn_Sprinkler_entry(P1);  // entry action
    _aCIP35_Conn_Sprinkler_active(N);  // step action
END_STEP
TRANSITION FROM CIP35_Conn_Sprinkler TO ReadyToCondition_Count
    := bStepDone;
END_TRANSITION
TRANSITION FROM Condition_CIP35_Client TO StopPump_CIP35_02
    := bCIP_Condition_Failed;
END_TRANSITION
STEP StopPump_CIP35_02:
    _aStopPump_CIP35_02_entry(P1);  // entry action
END_STEP
TRANSITION FROM StopPump_CIP35_02 TO ReFill_Water_T94
    := TRUE;
END_TRANSITION
STEP ReFill_Water_T94:
    _aReFill_Water_T94_active(N);  // step action
END_STEP
TRANSITION FROM ReFill_Water_T94 TO Condition_CIP35_Client
    := bStepDone;
END_TRANSITION
STEP Tank_LowLevel_CIP35_01:
    _aTank_LowLevel_CIP35_01_active(N);  // step action
END_STEP
TRANSITION FROM Tank_LowLevel_CIP35_01 TO CIP35_Done
    := bStepDone;
END_TRANSITION
STEP CIP35_Done:  // min time T#2s
    _aCIP35_Done_entry(P1);  // entry action
END_STEP
TRANSITION FROM CIP35_Done TO End_Check
    := TRUE;
END_TRANSITION
STEP End_Check:
    _aEnd_Check_active(N);  // step action
END_STEP
TRANSITION FROM End_Check TO Disconnect_n_Drain_CIP_Client
    := bStepDone;
END_TRANSITION
TRANSITION FROM End_Check TO Get_Client
    := TRUE;
END_TRANSITION
STEP Disconnect_n_Drain_CIP_Client:
    _aDisconnect_n_Drain_CIP_Client_entry(P1);  // entry action
    _aDisconnect_n_Drain_CIP_Client_active(N);  // step action
END_STEP
TRANSITION FROM Disconnect_n_Drain_CIP_Client TO Done
    := bStepDone;
END_TRANSITION
STEP Done:  // min time T#0.1s
    _aDone_entry(P1);  // entry action
END_STEP
TRANSITION FROM Done TO Disconnect_Old_Client
    := TRUE;
END_TRANSITION
// branch label Branch28_act_Oper
// branch label Branch29_act_Oper
// branch label Branch27_act_Oper
// branch label Branch26_act_Oper
// branch label Branch0_act_Oper
// branch label Branch11_act_Oper
// branch label Branch10_act_Oper
// branch label Branch15_act_Oper
// branch label Branch14_act_Oper
// branch label Branch10_act_Oper_2
// branch label Branch23_act_Oper
// branch label Branch12_act_Oper
// branch label Branch9_act_Oper
// branch label Branch17_act_Oper
// branch label Branch18_act_Oper
// branch label Branch19_act_Oper
// branch label Branch24_act_Oper
// branch label Branch20_act_Oper
// branch label Branch8_act_Oper
// branch label Branch2_act_Oper
// branch label Branch3_act_Oper
END_ACTION

ACTION act_ReqBuffer:
rtPosMoveHMI_Up(Q=>);
IF rtPosMoveHMI_Up.Q THEN;
	m_PosMove_Up_HMI();
END_IF
rtPosMoveHMI_Down(Q=>);
IF rtPosMoveHMI_Down.Q THEN;
	m_PosMove_Down_HMI();
END_IF
rtPosDeleteHMI(Q=>);
IF rtPosDeleteHMI.Q THEN;
	m_PosDelete_HMI();
END_IF
rtPosDeleteAllHMI(Q=>);
IF rtPosDeleteAllHMI.Q THEN;
	m_PosDeleteAll_HMI();
END_IF

rtReqLocalCIP_Full_HMI(Q=>);
IF rtReqLocalCIP_Full_HMI.Q THEN;
	eReqLocal.eClient:=E_CIP_Usage.eLocal;
	eReqLocal.eType:=E_CIP_Type.Full;
	m_TakePosInCIPBuffer(stCIP_Request:=eReqLocal);
END_IF

rtReqLocalCIP_Detergent_HMI(Q=>);
IF rtReqLocalCIP_Detergent_HMI.Q THEN;
	eReqLocal.eClient:=E_CIP_Usage.eLocal;
	eReqLocal.eType:=E_CIP_Type.Detergent;
	m_TakePosInCIPBuffer(stCIP_Request:=eReqLocal);
END_IF

rtReqCleanEmpty_HMI(Q=>);
IF rtReqCleanEmpty_HMI.Q THEN;
	m_CleanEmpty_Spaces();
END_IF
END_ACTION

ACTION act_Run:
//Client error: ALARM from Siemens. Only marks the step, the reaction is in FB_CIP_Siemens
IF eReq.eClient=E_CIP_Usage.eExternal THEN;
	IF g_Anybus.fbAnybus.stIn.bAlarm AND SFCCurrentStep<>'Ready' THEN;
		m_Set_LastStepBeforeError();
		sError_Message:='Client Error';
		//mResetCycle();
	END_IF
END_IF
END_ACTION

ACTION act_SprinklerCondition:


	IF TRUE
	AND eCIP_State>=E_Element_State_Long.eCIP_1_Rinzed 
	AND eCIP_State<=E_Element_State_Long.eCIP_2_Deterged 
	THEN;
		IF NOT bSprinkler THEN // Pipe
			tConditionTime	:=st_CIP_Param.t_ConditionDetergent;
			fFlowRate		:=st_CIP_Param.r_Flow_Pipe;
		ELSE // Sprinkler
			tConditionTime	:=st_CIP_Param.t_ConditionDetergent_Sprinkler;
			fFlowRate		:=st_CIP_Param.r_Flow_Sprinkler;
		END_IF	
		//rVolume_Collect :=st_CIP_Param.r_Volume_Collect_Detergent;
		//rVolume_Drain	:=st_CIP_Param.r_Volume_Drain_Detergent;
		//rVolume_Recycle	:=st_CIP_Param.r_Volume_Recycle_Detergent;
		
	ELSIF TRUE
	AND eCIP_State>=E_Element_State_Long.eCIP_3_Deterged_Clean 
	AND eCIP_State<=E_Element_State_Long.eCIP_4_Sanitized 
	THEN;
		IF NOT bSprinkler THEN // Pipe
			tConditionTime	:=st_CIP_Param.t_ConditionDisInfection;
			fFlowRate		:=st_CIP_Param.r_Flow_Pipe;
		ELSE // Sprinkler
			tConditionTime	:=st_CIP_Param.t_ConditionDisInfection_Sprinkler;
			fFlowRate		:=st_CIP_Param.r_Flow_Sprinkler;
		END_IF	
		//rVolume_Collect :=st_CIP_Param.r_Volume_Collect_DisInfection;
		//rVolume_Drain	:=st_CIP_Param.r_Volume_Drain_DisInfection;
		//rVolume_Recycle	:=st_CIP_Param.r_Volume_Recycle_DisInfection;
	END_IF
END_ACTION

METHOD m_Set_CIP_State : BOOL
VAR_INPUT
	eState	: E_Element_State_Long;
END_VAR
//CIP stages only move forward (eNotClean restarts)
IF (eState>eCIP_State
OR eState=E_Element_State_Long.eNotClean)
AND eState<=E_Element_State_Long.eProduction
THEN;
	eCIP_State:=eState;
	m_Set_CIP_State:=TRUE;
END_IF
END_METHOD

METHOD m_DashState_NotAvailable : BOOL
VAR_INPUT
	stage: E_CIP_DashStage_List;
END_VAR
//Client and sprinkler stages do not exist in the local CIP
CASE stage OF
	E_CIP_DashStage_List.e01_CIP1_Client_Drain_Product_Rest_Pipe,
	E_CIP_DashStage_List.e02_CIP1_Client_Drain_Product_Rest_Sprinkler,
	E_CIP_DashStage_List.e05_CIP2_Client_Detergent_Fill,
	E_CIP_DashStage_List.e06_CIP2_Client_Detergent_Condition_Pipe,
	E_CIP_DashStage_List.e07_CIP2_Client_Detergent_Condition_Sprinkler,
	E_CIP_DashStage_List.e11_CIP3_Detergent_Clean_Sprinkler,
	E_CIP_DashStage_List.e14_CIP4_Client_DisInfection_Fill,
	E_CIP_DashStage_List.e15_CIP4_Client_DisInfection_Condition_Pipe,
	E_CIP_DashStage_List.e16_CIP4_Client_DisInfection_Condition_Sprinkler,
	E_CIP_DashStage_List.e20_CIP5_DisInfection_Clean_Sprinkler:;
		m_DashState_NotAvailable:=TRUE;
ELSE;
		m_DashState_NotAvailable:=FALSE;
END_CASE
END_METHOD

METHOD m_Check_ProductionTank_Low_Level : BOOL
VAR_INPUT
END_VAR
//The client level is on the plant side: Tank waits for CLIENT EMPTY, as senLL before, Pipe passes
tonTankLowLevel.IN:=g_Anybus.fbAnybus.stIn.bClientEmpty;
tonTankLowLevel(PT:=T#2S);
IF bClientTypeIs_Tank
AND tonTankLowLevel.Q
THEN;
	m_Check_ProductionTank_Low_Level:=TRUE;
ELSIF NOT bClientTypeIs_Tank
THEN;
	m_Check_ProductionTank_Low_Level:=TRUE;
ELSE;
	m_Check_ProductionTank_Low_Level:=FALSE;
END_IF
END_METHOD

METHOD m_CleanEmpty_Spaces : BOOL
VAR_INPUT
END_VAR

VAR
	i: INT;
	j: INT;
	stCIP_Request_Empty: ST_CIP_Request;
END_VAR
FOR i:=0 TO 9 DO
	IF i<>0 OR NOT bRun THEN;
		IF arCIP_RequestBufer[i].eClient=E_CIP_Usage.eNotInUse THEN;
			FOR j:=i+1 TO 9 DO
				IF arCIP_RequestBufer[j].eClient<>E_CIP_Usage.eNotInUse THEN;
					arCIP_RequestBufer[i]:=arCIP_RequestBufer[j];
					arCIP_RequestBufer[j]:=stCIP_Request_Empty;
					EXIT;
				END_IF
			END_FOR
		END_IF		
	END_IF
END_FOR
END_METHOD

METHOD m_ClientTank_IsEmpty : BOOL
VAR_INPUT
END_VAR
IF __ISVALIDREF(ref_lvlTank_Client) 
AND bClientTypeIs_Tank
THEN;
	m_ClientTank_IsEmpty:=ref_lvlTank_Client.e_state=E_Tank_Level.eEmpty;
ELSE;
	m_ClientTank_IsEmpty:=TRUE;
END_IF
END_METHOD

METHOD m_ClientTank_Level_IsHigher_Then : BOOL
VAR_INPUT
	min_Level: REAL:=150.0;
END_VAR
IF __ISVALIDREF(ref_lvlTank_Client) 
AND bClientTypeIs_Tank
THEN;
	m_ClientTank_Level_IsHigher_Then:=ref_lvlTank_Client.rTankLevel>=min_Level;
ELSE;
	m_ClientTank_Level_IsHigher_Then:=FALSE;
END_IF
END_METHOD

METHOD m_DashState_activate : BOOL
VAR_INPUT
	stage		: E_CIP_DashStage_List;
END_VAR
	IF arCIP_DashStage_list[stage] = E_CIP_DashStage.eCIPStage_ToBeDone THEN;
		arCIP_DashStage_list[stage]:=E_CIP_DashStage.eCIPStage_Active;
		eCIP_DashStage_actual:=stage;
		sCIP_DashStage_actual:=TO_STRING(eCIP_DashStage_actual);	
		RETURN;
	END_IF

(*
FOR stage:=m_DashState_from() TO m_DashState_to() DO
	IF arCIP_DashStage_list[stage] = E_CIP_DashStage.eCIPStage_ToBeDone THEN;
		arCIP_DashStage_list[stage]:=E_CIP_DashStage.eCIPStage_Active;
		eCIP_DashStage_actual:=stage;
		sCIP_DashStage_actual:=TO_STRING(eCIP_DashStage_actual);	
		RETURN;
	END_IF
END_FOR
*)
END_METHOD

METHOD m_DashState_done : BOOL
VAR_INPUT
	stage	: E_CIP_DashStage_List;
END_VAR
IF arCIP_DashStage_list[stage] = E_CIP_DashStage.eCIPStage_Active THEN;
	arCIP_DashStage_list[stage]:=E_CIP_DashStage.eCIPStage_Done;
	RETURN;
END_IF

(*
FOR stage:=m_DashState_from() TO m_DashState_to() DO
	IF arCIP_DashStage_list[stage] = E_CIP_DashStage.eCIPStage_Active THEN;
		arCIP_DashStage_list[stage]:=E_CIP_DashStage.eCIPStage_Done;
		RETURN;
	END_IF
END_FOR
*)
END_METHOD

METHOD m_DashState_from : E_CIP_DashStage_List
VAR
	eActCIP_State	: E_Element_State_Long;
END_VAR
eActCIP_State:=eCIP_State;

CASE eActCIP_State OF
	E_Element_State_Long.eNotClean:;
		m_DashState_from:=E_CIP_DashStage_List.e01_CIP1_Client_Drain_Product_Rest_Pipe;	
		
	E_Element_State_Long.eCIP_1_Rinzed:;
		m_DashState_from:=E_CIP_DashStage_List.e03_CIP2_Local_Detergent_Fill;	
	
	E_Element_State_Long.eCIP_2_Deterged:;
		m_DashState_from:=E_CIP_DashStage_List.e08_CIP3_Detergent_Collect;	
	
	E_Element_State_Long.eCIP_3_Deterged_Clean:;
		m_DashState_from:=E_CIP_DashStage_List.e12_CIP4_Local_DisInfection_Fill;	
	
	E_Element_State_Long.eCIP_4_Sanitized:;
		m_DashState_from:=E_CIP_DashStage_List.e17_CIP5_DisInfection_Collect;	
	
ELSE;
	//???
		m_DashState_from:=E_CIP_DashStage_List.eLast;
END_CASE
END_METHOD

METHOD m_DashState_Get_ToBeDone_List : BOOL
VAR
	//eActCIP_State	: E_Element_State_Long;
	//eCIP_req		: ST_CIP_Request;	
	stage			: E_CIP_DashStage_List;
END_VAR
//eCIP_req:=eReq;

//init
FOR stage:=E_CIP_DashStage_List.e00_NotSelected TO E_CIP_DashStage_List.eLast DO
	arCIP_DashStage_list[stage]:=E_CIP_DashStage.eCIPStage_NotAvalable;
END_FOR

//Start done condition stages
FOR stage:=E_CIP_DashStage_List.e00_NotSelected TO m_DashState_from()-1 DO
	IF m_DashState_Sprinkler(stage:=stage) THEN;
		IF bClientTypeIs_Tank THEN;
			arCIP_DashStage_list[stage]:=E_CIP_DashStage.eCIPStage_Done;
		ELSE;
			arCIP_DashStage_list[stage]:=E_CIP_DashStage.eCIPStage_NotAvalable;
		END_IF
	ELSE;
		arCIP_DashStage_list[stage]:=E_CIP_DashStage.eCIPStage_Done;
	END_IF
END_FOR

// Request conditions
FOR stage:=m_DashState_from() TO m_DashState_to() DO
	IF m_DashState_Sprinkler(stage:=stage) THEN;
		IF bClientTypeIs_Tank THEN;
			arCIP_DashStage_list[stage]:=E_CIP_DashStage.eCIPStage_ToBeDone;
		ELSE;
			arCIP_DashStage_list[stage]:=E_CIP_DashStage.eCIPStage_NotAvalable;
		END_IF
	ELSE;
		arCIP_DashStage_list[stage]:=E_CIP_DashStage.eCIPStage_ToBeDone;
	END_IF
END_FOR

//Do not requested 
FOR stage:=m_DashState_to()+1 TO E_CIP_DashStage_List.eLast DO
	IF m_DashState_Sprinkler(stage:=stage) THEN;
		IF bClientTypeIs_Tank THEN;
			arCIP_DashStage_list[stage]:=E_CIP_DashStage.eCIPStage_NotInUse;
		ELSE;
			arCIP_DashStage_list[stage]:=E_CIP_DashStage.eCIPStage_NotAvalable;
		END_IF
	ELSE;
		arCIP_DashStage_list[stage]:=E_CIP_DashStage.eCIPStage_NotInUse;
	END_IF
END_FOR
END_METHOD

METHOD m_DashState_Sprinkler : BOOL
VAR_INPUT
	stage: E_CIP_DashStage_List;
END_VAR
CASE stage OF 
	E_CIP_DashStage_List.e02_CIP1_Client_Drain_Product_Rest_Sprinkler,
	E_CIP_DashStage_List.e07_CIP2_Client_Detergent_Condition_Sprinkler,
	E_CIP_DashStage_List.e11_CIP3_Detergent_Clean_Sprinkler,
	E_CIP_DashStage_List.e16_CIP4_Client_DisInfection_Condition_Sprinkler,
	E_CIP_DashStage_List.e20_CIP5_DisInfection_Clean_Sprinkler:;
		m_DashState_Sprinkler:=TRUE;
ELSE;
		m_DashState_Sprinkler:=FALSE;
END_CASE
END_METHOD

METHOD m_DashState_to : E_CIP_DashStage_List
VAR
	eCIP_req		: ST_CIP_Request;
END_VAR
eCIP_req:=eReq;

CASE eCIP_req.eType OF
	E_CIP_Type.R_Water:;
		m_DashState_to:=E_CIP_DashStage_List.e02_CIP1_Client_Drain_Product_Rest_Sprinkler;
		
	E_CIP_Type.Detergent:;
		m_DashState_to:=E_CIP_DashStage_List.e11_CIP3_Detergent_Clean_Sprinkler;
	
	E_CIP_Type.Full:;
		m_DashState_to:=E_CIP_DashStage_List.e20_CIP5_DisInfection_Clean_Sprinkler;

ELSE;
	//???
		m_DashState_to:=E_CIP_DashStage_List.eLast;	
END_CASE
END_METHOD

METHOD m_DashState_ToString_convertion : BOOL
VAR_INPUT
END_VAR

VAR
	eDashboard_CIP_State: E_CIP_DashStage_List:=E_CIP_DashStage_List.eLast;
END_VAR
FOR eDashboard_CIP_State:=0 TO E_CIP_DashStage_List.eLast DO
	//g_HMI.arCIP_DashStage_list[eDashboard_CIP_State]:=E_CIP_DashStage.eCIPStage_NotInUse;
	g_HMI.arCIP_DashStage_string[eDashboard_CIP_State]:=TO_STRING(eDashboard_CIP_State);
END_FOR
END_METHOD

METHOD m_MeasureTimeToHMI : TIME
VAR_INPUT
END_VAR
IF SFCCurrentStep='measureDelay_CIP2_1' THEN;
	m_MeasureTimeToHMI:=measureDelay_CIP2_1.t;
	
ELSIF SFCCurrentStep='measureDelay_CIP2_2' THEN;
	m_MeasureTimeToHMI:=measureDelay_CIP2_2.t;
	
ELSIF SFCCurrentStep='measureDelay_CIP4_1' THEN;
	m_MeasureTimeToHMI:=measureDelay_CIP4_1.t;
	
ELSIF SFCCurrentStep='measureDelay_CIP4_2' THEN;
	m_MeasureTimeToHMI:=measureDelay_CIP4_2.t;

ELSE;
	m_MeasureTimeToHMI:=T#0S;
END_IF
END_METHOD

METHOD m_OverFlowCorrect : REAL
VAR_INPUT
	rTc		:	REAL	;//Target concentration
	rAv		:	REAL	;//Actual volume
	rAc		:	REAL	;//Actual concentration
END_VAR
//Calculating the additional valume of fresh water to dalute the concentration
IF rTc=0 THEN;
	m_OverFlowCorrect:=0;
ELSE;
	m_OverFlowCorrect:=((rAv*rAc/100)/(rTc/100))-(rAv*rAc/100)-rAv+(rAv*rAc/100);
END_IF
END_METHOD

METHOD m_PosDelete_HMI : BOOL
VAR_INPUT
END_VAR
VAR
	stCIP_Request_Empty: ST_CIP_Request;
END_VAR
IF iPosSelect_HMI>=0 AND iPosSelect_HMI<9 THEN;
	IF iPosSelect_HMI<>0 OR NOT bRun THEN;
		arCIP_RequestBufer[iPosSelect_HMI]:=stCIP_Request_Empty;
	END_IF		
END_IF
END_METHOD

METHOD m_PosDeleteAll_HMI : BOOL
VAR_INPUT
END_VAR
VAR
	stCIP_Request_Empty: ST_CIP_Request;
	i: INT;
END_VAR

FOR i:=0 TO 9 DO
	IF i<>0 OR NOT bRun THEN;
		arCIP_RequestBufer[i]:=stCIP_Request_Empty;
	END_IF	
END_FOR
END_METHOD

METHOD m_PosMove_Down_HMI : BOOL
VAR_INPUT
END_VAR
VAR
	stCIP_Request_Temp: ST_CIP_Request;
	i: INT;
END_VAR
IF iPosSelect_HMI>=0 AND iPosSelect_HMI<9 THEN;
	IF iPosSelect_HMI<>0 OR NOT bRun THEN;		
			IF ((arCIP_RequestBufer[iPosSelect_HMI].eType=E_CIP_Type.R_Water 
				AND (arCIP_RequestBufer[iPosSelect_HMI+1].eType=E_CIP_Type.Detergent 
				OR arCIP_RequestBufer[iPosSelect_HMI+1].eType=E_CIP_Type.Full)) 
			OR (arCIP_RequestBufer[iPosSelect_HMI].eType=E_CIP_Type.Detergent 				
				AND arCIP_RequestBufer[iPosSelect_HMI+1].eType=E_CIP_Type.Full))
			AND (arCIP_RequestBufer[iPosSelect_HMI+1].eClient=arCIP_RequestBufer[iPosSelect_HMI].eClient) 
			THEN
				;
			ELSE
				stCIP_Request_Temp:=arCIP_RequestBufer[iPosSelect_HMI+1];
				arCIP_RequestBufer[iPosSelect_HMI+1]:=arCIP_RequestBufer[iPosSelect_HMI];
				arCIP_RequestBufer[iPosSelect_HMI]:=stCIP_Request_Temp;
				iPosSelect_HMI:=iPosSelect_HMI+1;	
			END_IF	
	END_IF
END_IF
END_METHOD

METHOD m_PosMove_Up_HMI : BOOL
VAR_INPUT
END_VAR
VAR
	stCIP_Request_Temp: ST_CIP_Request;
	i: INT;
	m: bool;
END_VAR
IF iPosSelect_HMI>0 AND iPosSelect_HMI<=9 THEN;
	IF iPosSelect_HMI<>1 OR NOT bRun THEN;			
			IF ((arCIP_RequestBufer[iPosSelect_HMI].eType=e_cip_type.Full 
				AND (arCIP_RequestBufer[iPosSelect_HMI-1].eType=E_CIP_Type.Detergent 
				OR arCIP_RequestBufer[iPosSelect_HMI-1].eType=E_CIP_Type.R_Water)) 
			OR (arCIP_RequestBufer[iPosSelect_HMI].eType=E_CIP_Type.Detergent 
				AND arCIP_RequestBufer[iPosSelect_HMI-1].eType=E_CIP_Type.R_Water))
			AND (arCIP_RequestBufer[iPosSelect_HMI-1].eClient=arCIP_RequestBufer[iPosSelect_HMI].eClient) 
			THEN
				;
			ELSE
				stCIP_Request_Temp:=arCIP_RequestBufer[iPosSelect_HMI-1];
				arCIP_RequestBufer[iPosSelect_HMI-1]:=arCIP_RequestBufer[iPosSelect_HMI];
				arCIP_RequestBufer[iPosSelect_HMI]:=stCIP_Request_Temp;
				iPosSelect_HMI:=iPosSelect_HMI-1;
			END_IF	
	END_IF
END_IF
END_METHOD

METHOD m_Set_SFCFlags_Reference : BOOL
//Set reference to SFC flags

refSFC.SFCInit REF= SFCInit;
refSFC.SFCReset REF= SFCReset;
refSFC.SFCError REF= SFCError;
refSFC.SFCEnableLimit REF= SFCEnableLimit;
refSFC.SFCErrorStep REF= SFCErrorStep;
refSFC.SFCErrorPOU REF= SFCErrorPOU;
refSFC.SFCQuitError REF= SFCQuitError;
refSFC.SFCPause REF= SFCPause;
refSFC.SFCTrans REF= SFCTrans;
refSFC.SFCCurrentStep REF= SFCCurrentStep;
refSFC.SFCTip REF= SFCTip;
refSFC.SFCTipMode REF= SFCTipMode;

// Cycle handle for SFC
m_SFC_Handle();

m_Set_Mode_Reference(inMoedeZone:=E_ModeZone.eCIP);
END_METHOD

METHOD m_TakePosInCIPBuffer : BOOL
VAR_INPUT
	stCIP_Request: ST_CIP_Request;
END_VAR

VAR
	i: INT;
	m: bool;	
END_VAR
//Old client checks (production, state, duplicate), not used for eExternal, fbElement is removed
(*
IF stCIP_Request.eClient<>E_CIP_Usage.eNotInUse
AND stCIP_Request.eType<>E_CIP_Type.NotSelected
AND g_data.fbElement[stCIP_Request.eClient].ProdStatus<>E_Prod_Status.Active
AND g_data.fbElement[stCIP_Request.eClient].eState_Long>E_Element_State_Long.eStandby 
AND ((stCIP_Request.eType=E_CIP_Type.R_Water AND g_data.fbElement[stCIP_Request.eClient].eState_Long<E_Element_State_Long.eCIP_1_Rinzed)
	OR (stCIP_Request.eType=E_CIP_Type.Detergent AND g_data.fbElement[stCIP_Request.eClient].eState_Long<E_Element_State_Long.eCIP_3_Deterged_Clean)
	OR (stCIP_Request.eType=E_CIP_Type.Full AND g_data.fbElement[stCIP_Request.eClient].eState_Long<E_Element_State_Long.eCIP_5_Done))

THEN
	FOR i:=0 TO 9 DO
		IF arCIP_RequestBufer[i].eClient=stCIP_Request.eClient 
			AND arCIP_RequestBufer[i].eType>=stCIP_Request.eType 
		THEN 	
				m:=FALSE;
				EXIT;
			ELSE
				m:=TRUE;
		END_IF
	END_FOR	
	IF m=TRUE THEN
		FOR i:=0 TO 9 DO
			IF arCIP_RequestBufer[i].eClient=E_CIP_Usage.eNotInUse 
			THEN;
				arCIP_RequestBufer[i]:=stCIP_Request;
				m:=FALSE;
				EXIT;
			END_IF
		END_FOR	
	END_IF
ELSIF stCIP_Request.eClient=E_CIP_Usage.eLocal
AND stCIP_Request.eType<>E_CIP_Type.NotSelected
THEN;
		FOR i:=0 TO 9 DO
			IF arCIP_RequestBufer[i].eClient=E_CIP_Usage.eNotInUse 
			THEN;
				arCIP_RequestBufer[i]:=stCIP_Request;
				m:=FALSE;
				EXIT;
			END_IF
		END_FOR		
END_IF
*)
//R_Water is not a valid local request
IF (stCIP_Request.eClient=E_CIP_Usage.eLocal
	AND (stCIP_Request.eType=E_CIP_Type.Detergent OR stCIP_Request.eType=E_CIP_Type.Full))
OR (stCIP_Request.eClient=E_CIP_Usage.eExternal
	AND stCIP_Request.eType<>E_CIP_Type.NotSelected)
THEN;
		FOR i:=0 TO 9 DO
			IF arCIP_RequestBufer[i].eClient=E_CIP_Usage.eNotInUse
			THEN;
				arCIP_RequestBufer[i]:=stCIP_Request;
				m:=FALSE;
				EXIT;
			END_IF
		END_FOR
END_IF
END_METHOD

METHOD mFillWater : BOOL
VAR_INPUT
END_VAR

VAR
	reqVolume: REAL;	
	valve : E_Pis_Name;;
	actLevel: REAL;
	fillCondition: BOOL;	
	
END_VAR
IF TRUE 
AND fbPis.m_CheckByRecipe(stPis:=stPis_FillWater_T91, req:=E_Piston_Recipe_State.Release)
AND fbPis.m_CheckByRecipe(stPis:=stPis_FillWater_T92, req:=E_Piston_Recipe_State.Release)
AND fbPis.m_CheckByRecipe(stPis:=stPis_FillWater_T93, req:=E_Piston_Recipe_State.Release)
AND bStateSafe
AND MAIN.bTemp_Water_Overweight_check
THEN;
	fillCondition:=TRUE;
ELSE;
	fillCondition:=FALSE;
END_IF

reqVolume:=st_CIP_Param.r_Tank94_Volume;
IF g_Data.arr_CIP_Recipe[nLocalRecipe].r_Tank94_Volume>reqVolume THEN;
	reqVolume:=g_Data.arr_CIP_Recipe[nLocalRecipe].r_Tank94_Volume;
END_IF

fbHysteresisFillT94(
	fIn:= lvlTank_T94.rTankLevel, 
	fHigh:= reqVolume, 
	fLow:= reqVolume-50.0, 
	iDigitsAfterDot:= 1, 
	bOut=> );

IF eMode<>E_CIP_Mode.eOff THEN;
	IF fbPis.m_CheckByRecipe(stPis:=stPis_FillWater_T94, req:=E_Piston_Recipe_State.Act) 
	AND (NOT fbHysteresisFillT94.bOut
	OR NOT fillCondition)
	THEN;
		//stPis_FillWater_T94.req_Close:=TRUE;
		fbPis.m_SetByRecipe(stPis:=stPis_FillWater_T94, req:=E_Piston_Recipe_State.Release);
		
	ELSIF fbPis.m_CheckByRecipe(stPis:=stPis_FillWater_T94, req:=E_Piston_Recipe_State.Release) 
	AND fbHysteresisFillT94.bOut
	AND fillCondition
	THEN;
		IF NOT arrTanksSens[E_Tank_Name.T94].get_stTankLevel_OverFlow() THEN;
			fbPis.m_SetByRecipe(stPis:=stPis_FillWater_T94, req:=E_Piston_Recipe_State.Act);			
		END_IF	
	END_IF	
END_IF
	
	
(*
fbFillT94(	
		valve:= valFillWater_T94, 
		reqLevel:= reqVolume, 
		actLevel:= lvlTank_T94.rTankLevel, 
		fillCondition:= );
*)
END_METHOD

METHOD mLoadDefProcessSetPoints : BOOL
VAR_INPUT
END_VAR

	stDetergent.ToleranceHigh:=0.05;
	stDetergent.ToleravceLow:=0.05;
	stTemperature_Deterg.ToleranceHigh:=1;
	stTemperature_Deterg.ToleravceLow:=1;
	stDisInfectant.ToleranceHigh:=0.05;
	stDisInfectant.ToleravceLow:=0.05;
	stTemperature_Dis.ToleranceHigh:=1;//0.5
	stTemperature_Dis.ToleravceLow:=1;//0.5
	stFlow1_Rate.ToleranceHigh:=10;
	stFlow1_Rate.ToleravceLow:=10;
	stFlow2_Rate.ToleranceHigh:=10;
	stFlow2_Rate.ToleravceLow:=10;
	stP1001_Pressure.ToleranceHigh:=1;
	stP1001_Pressure.ToleravceLow:=1;
END_METHOD

METHOD mProcessDeviation : REAL
VAR_INPUT
	reqValue: REAL;
	processValue: REAL;
END_VAR
mProcessDeviation:=reqValue-processValue;
END_METHOD

METHOD mVolumeMeter : BOOL
VAR_INPUT
END_VAR
delta_T91_Volume:=lvlTank_T91.rTankLevel-memo_T91_Level_start;//de
delta_T92_Volume:=lvlTank_T92.rTankLevel-memo_T92_Level_start;
delta_T93_Volume:=lvlTank_T93.rTankLevel-memo_T93_Level_start;
delta_T94_Volume:=lvlTank_T94.rTankLevel-memo_T94_Level_start;
END_METHOD

METHOD mVolumeReset_All : BOOL
VAR_INPUT
END_VAR
memo_T91_Level_start:=lvlTank_T91.rTankLevel;
memo_T92_Level_start:=lvlTank_T92.rTankLevel;
memo_T93_Level_start:=lvlTank_T93.rTankLevel;
memo_T94_Level_start:=lvlTank_T94.rTankLevel;
END_METHOD

END_FUNCTION_BLOCK

// ---- 00 Library/13 Process Control/FB_ProcessControl.TcPOU
FUNCTION_BLOCK FB_ProcessControl

VAR_IN_OUT
	stProcessControl	:	ST_ProcessControl	;
END_VAR
VAR
	bRun			: BOOL	;
	//fbPID	: 	FB_BasicPID	;
	fbPID	: 	PID	;
	hystCIP_SetPoint: FB_Hysteresis_REAL;
	Call_ActDelayTON	: TON	;
	bRunCalled		: BOOL	;//mRun was called since the last body call

	handling_PID_Manual: TON;

END_VAR

//stProcessControl.bManual:=TRUE;



//Deactivate control 1s after mRun stops being called (body may be called several times per cycle)
Call_ActDelayTON(IN:=stProcessControl.bActiveCntr AND NOT bRunCalled , PT:=T#1S , Q=> , ET=> );
bRunCalled:=FALSE;

m_Check();

act_Call_PID();
act_CallHyst();

handling_PID_Manual(PT:=T#0.5S);//, IN:=TRUE
IF handling_PID_Manual.Q THEN;
	stProcessControl.bManual:=TRUE;
ELSE;
	stProcessControl.bManual:=FALSE;
END_IF

ACTION act_Call_PID:
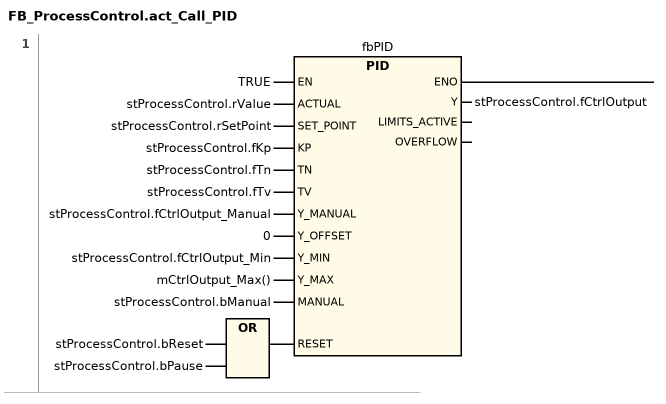
// NETWORK 1
fbPID(
    ACTUAL := stProcessControl.rValue,
    SET_POINT := stProcessControl.rSetPoint,
    KP := stProcessControl.fKp,
    TN := stProcessControl.fTn,
    TV := stProcessControl.fTv,
    Y_MANUAL := stProcessControl.fCtrlOutput_Manual,
    Y_OFFSET := 0,
    Y_MIN := stProcessControl.fCtrlOutput_Min,
    Y_MAX := mCtrlOutput_Max(),
    MANUAL := stProcessControl.bManual,
    RESET := stProcessControl.bReset OR stProcessControl.bPause,
    Y => stProcessControl.fCtrlOutput); // PID
END_ACTION

ACTION act_Call_PID_old:

	
(*
fbPID(
	fSetpointValue:=stProcessControl.rSetPoint , 
	fActualValue:=stProcessControl.rValue , 
	bReset:=stProcessControl.bReset , 
	fCtrlCycleTime:=stProcessControl.fCtrlCycleTime , 
	fKp:=stProcessControl.fKp , 
	fTn:=stProcessControl.fTn , 
	fTv:=stProcessControl.fTv , 
	fTd:=stProcessControl.fTd , 
	fCtrlOutput=>stProcessControl.fCtrlOutput , 
	nErrorStatus=>stProcessControl.nErrorStatus );
*)
END_ACTION

ACTION act_CallHyst:
hystCIP_SetPoint(
	fIn:=stProcessControl.rValue,//g_HMI.stT4_Sens.rTankLevel,
	fHigh:=stProcessControl.fHystHigh,
	fLow:=stProcessControl.fHystLow,
	iDigitsAfterDot:=,
	bOut=>stProcessControl.bHystOut);
END_ACTION

METHOD m_Check : BOOL
VAR_INPUT
END_VAR
IF NOT __ISVALIDREF(stProcessControl) THEN
	RETURN;
END_IF

IF bRun THEN
	stProcessControl.bActiveCntr:=TRUE;
	bRunCalled:=TRUE;
ELSIF NOT bRun AND Call_ActDelayTON.Q THEN
	stProcessControl.bActiveCntr:=FALSE;
END_IF

IF bRun THEN
	stProcessControl.Deviation:=stProcessControl.rSetPoint-stProcessControl.rValue;
	stProcessControl.Control_ON:=FALSE;
	stProcessControl.OverFlow:=FALSE;
	stProcessControl.bDone:=FALSE;
	
	IF stProcessControl.Deviation >= stProcessControl.ToleravceLow THEN;
		//Value too low needs to be increased
		stProcessControl.Control_ON:=TRUE;
		stProcessControl.OverFlow:=FALSE;
		stProcessControl.bDone:=FALSE;
	ELSIF stProcessControl.Deviation <= -stProcessControl.ToleranceHigh THEN;
		//value too high need to be decreased
		stProcessControl.OverFlow:=TRUE;
		stProcessControl.Control_ON:=TRUE;
		stProcessControl.bDone:=FALSE;
		//message
	ELSE;
		// Done, value in tolerace
		stProcessControl.OverFlow:=FALSE;
		stProcessControl.Control_ON:=FALSE;
		stProcessControl.bDone:=TRUE;
	END_IF
	bRun:=FALSE;
END_IF
END_METHOD

METHOD mCtrlOutput_Max : REAL
VAR_INPUT
END_VAR

VAR
	span: LREAL;
END_VAR


span:=ABS(stProcessControl.fCtrlOutput_Max-stProcessControl.fCtrlOutput_Min);
//LimitedPrecentage:=
IF stProcessControl.rValue>stProcessControl.rValue_Min_To_ReleaseControl THEN;
	mCtrlOutput_Max:=stProcessControl.fCtrlOutput_Max;
ELSE;
	mCtrlOutput_Max:=stProcessControl.fCtrlOutput_Min+(span*0.3);
END_IF
END_METHOD

METHOD mManual : BOOL
VAR_INPUT
	value: BOOL;
END_VAR
//PID manual request without starting control (bRun/bActiveCntr untouched)
handling_PID_Manual(IN:=value);
mManual:=stProcessControl.bManual;
END_METHOD

METHOD mPause : BOOL
VAR_INPUT
	value: BOOL;
END_VAR
stProcessControl.bPause:=value;
END_METHOD

METHOD mReset : BOOL
VAR_INPUT
END_VAR
stProcessControl.Control_ON:=FALSE;
stProcessControl.OverFlow:=FALSE;
stProcessControl.bDone:=FALSE;
END_METHOD

METHOD mRun : BOOL
VAR_INPUT
	//Set_Point: REAL;
END_VAR
bRun:=TRUE;
//stProcessControl.rSetPoint:=Set_Point;
m_Check();



mRun:=stProcessControl.bDone;
END_METHOD

METHOD mRun_Hyst : REAL
VAR_INPUT
END_VAR
stProcessControl.bManual:=FALSE;
IF stProcessControl.bHystOut THEN
	mRun_Hyst:=stProcessControl.rHystOutLow;
ELSE
	mRun_Hyst:=stProcessControl.rHystOutHigh;
END_IF
END_METHOD

METHOD mRun_PID : REAL
VAR_INPUT
	Set_Point: REAL;
	controlManual: BOOL;
END_VAR
mRun();//mRun(Set_Point:=Set_Point);
//stProcessControl.bManual:=controlManual;
//stProcessControl.rSetPoint:=Set_Point;
handling_PID_Manual(IN:=controlManual);
mRun_PID:=stProcessControl.fCtrlOutput;
END_METHOD

METHOD mRun_With_SP : BOOL
VAR_INPUT
	Set_Point: REAL;
END_VAR
stProcessControl.rSetPoint:=Set_Point;
bRun:=TRUE;
mRun();
//stProcessControl.rSetPoint:=Set_Point;
mRun_With_SP:=stProcessControl.bDone;
END_METHOD

END_FUNCTION_BLOCK

// ---- 00 Library/10 Utils/FB_Hysteresis_REAL.TcPOU
FUNCTION_BLOCK FB_Hysteresis_REAL
VAR_INPUT
	fIn		: REAL; // in case of iDigitsAfterDot=2 max value 327.67 * 100 >> INTEGER Value limitation
	fHigh	: REAL;
	fLow	: REAL;
	iDigitsAfterDot: INT:=1; //min 0 , max 3

END_VAR
VAR_OUTPUT
	bOut	: BOOL;
END_VAR
VAR
	fbHys: HYSTERESIS;
	mult: INT;
	iDigitsAfterDot_Local: INT:=2; //min 0 , max 3


END_VAR

IF iDigitsAfterDot < 0 THEN;
	iDigitsAfterDot_Local:=0;
ELSIF iDigitsAfterDot > 3 THEN;
	iDigitsAfterDot_Local:=3;
ELSE;
	iDigitsAfterDot_Local:=iDigitsAfterDot;
END_IF
 

CASE iDigitsAfterDot_Local OF
	0:mult:=1;
	1:mult:=10;
	2:mult:=100;
	3:mult:=1000;
END_CASE

fbHys.HIGH:=REAL_TO_INT(fHigh*mult);
fbHys.LOW:=REAL_TO_INT(fLow*mult);
fbHys.IN:=REAL_TO_INT(fIn*mult);

fbHys(OUT=>bOut);

END_FUNCTION_BLOCK

// ---- 00 Library/10 Utils/TONR.TcPOU
FUNCTION_BLOCK TONR //Retentive Timer
VAR_INPUT
    IN : BOOL;         // Input signal
	ResetTime: BOOL;	//Reset Accumulating Time
    PT : TIME := T#0S; // Preset time
END_VAR
VAR_OUTPUT
    Q : BOOL;          // Output signal (true when time is reached)
    ET : TIME;         // Elapsed time
END_VAR
VAR
    StartTime : TIME := T#0S; // Start time storage
    IsTiming : BOOL := FALSE; // Timing state
END_VAR

// Start or continue timing when the input is true
IF IN THEN
    IF NOT IsTiming THEN
        StartTime := DT_TO_TIME(dtRealTime) - ET; // Adjust start time if resuming
        IsTiming := TRUE;
    END_IF
    ET := DT_TO_TIME(dtRealTime) - StartTime; // Calculate elapsed time
ELSE
    IsTiming := FALSE; // Stop timing but retain elapsed time
END_IF

IF ResetTime THEN
	ResetTime:=FALSE;
	IsTiming := FALSE; // Stop timing but retain elapsed time
	ET:=T#0s;
END_IF
 
// Check if the elapsed time has reached the preset time
IF ET >= PT THEN
    Q := TRUE;
ELSE
    Q := FALSE;
END_IF

END_FUNCTION_BLOCK

// ---- 00 Library/02 Pump/FB_Pump.TcPOU
FUNCTION_BLOCK FB_Pump
VAR_INPUT
	Pump_ID				: E_Pump_List:=E_Pump_List.eNotSelected;
	PressureSensor_ID	: E_ASense_Name:=E_ASense_Name.eNotSelected;
END_VAR
VAR
	sID: STRING(6);

	stNidec: REFERENCE TO ST_Nidec;
	status_word: WORD;
	control_word: WORD;

	ControlWord: ControlWordStruct;
	StatusWord: StatusWordStruct;


	//request
	modeAuto	:	BOOL	:= TRUE	;//System in automatic
	bRun_Auto	:	BOOL	;
	bRun_Man	:	BOOL	;

	//nRPM_Auto	:	REAL		;//Pump RPM 
	//nRPM_Man	:	REAL		;//Pump RPM 
	//feedback
	nRPM_fdbk	:	INT	;	
	rtManual: R_TRIG;
	ton_Drive_init: TON;
	state_init: (OFF,stage1,stage2,stage3,stage4, Ready);

	bInitiated: BOOL;
	ton_RPM_feedback_lag_monitoring: TON;
	ton_Pressure_feedback_monitoring: TON;
	
	fbPressureSensor: REFERENCE TO FB_AnalogSensor;

END_VAR
VAR_OUTPUT
	DriveReady	:   BOOL;
	bRun		: 	BOOL;
	nRPM		:	REAL		;//Pump RPM 
	
END_VAR
VAR_IN_OUT
	stPump			: ST_Pump	;
	stOperation		: ST_OperationButtons;
END_VAR

stNidec REF= gIO.Nidec[Pump_ID];
sID:=TO_STRING(Pump_ID);
nRPM:=stPump.nRPM;
IF __ISVALIDREF(stNidec) THEN;
	//run
	status_word:=stNidec.StatusWord;
	stNidec.ControlWord:=control_word;
	
	control_word:=m_Map_ControlWord(cwStruct:=ControlWord);
	StatusWord:=m_Map_StatusWord(wordInput:=status_word);
	
	stNidec.targetVelocity:=DINT_TO_INT(TRUNC(stPump.nRPM));	
	nRPM_fdbk:=stNidec.actVelocity;	
	
	m_Nidec_Init();
	
	IF state_init=Ready THEN;
		DriveReady:=TRUE;
		ControlWord.EnableOperation:=bRun;
	ELSE;
		DriveReady:=FALSE;
		//bRun:=bRun_Man:=bRun_Auto:=FALSE;
		ControlWord.EnableOperation:=FALSE;
	END_IF	
	stPump.DriveReady:=DriveReady;
ELSE;
	//RETURN;
END_IF

IF modeAuto THEN;
	//bRun:=bRun_Auto;
	IF bRun_Auto AND m_CheckOper() THEN;
		bRun:=TRUE;
	ELSE;
		bRun:=FALSE;
	END_IF
	stPump.nRPM:=stPump.nRPM_Auto;
ELSE;
	//bRun:=bRun_Man;
	IF bRun_Man AND m_CheckOper() THEN;
		bRun:=TRUE;
	ELSE;
		bRun:=FALSE;
	END_IF	
	stPump.nRPM:=stPump.nRPM_Man;
END_IF

rtManual(CLK:=NOT modeAuto);
IF rtManual.Q THEN;
	bRun:=bRun_Man:=bRun_Auto;
	//stPump.nRPM:=stPump.nRPM_Man:=stPump.nRPM_Auto;
END_IF

IF stPump.nRPM>3000 THEN;
	stPump.nRPM:=3000;
END_IF

stPump.bRun_Man:=bRun_Man;
stPump.bRun_Auto:=bRun_Auto;
stPump.bRun:=bRun;

IF m_Error()<>'' THEN;
	//stOperation.bSetPause:=TRUE;
	//print error
	//fbPrintErrMessageByID(sModuleDescription:='Pump',sActErrorID:='101x000x001');	
END_IF

bInitiated:=TRUE;

METHOD m_Auto : BOOL
VAR_INPUT
	control: LREAL; // RPM
END_VAR

VAR
	RPM: INT;
END_VAR
//ST_Pump.bRun_Auto:=TRUE;
m_Auto:=TRUE;
RPM:=DINT_TO_INT(TRUNC(control));
IF RPM>3000 THEN;
	stPump.nRPM_Auto:=3000;
ELSIF RPM<200 THEN;
	stPump.nRPM_Auto:=200;
ELSE;
	stPump.nRPM_Auto:=RPM;
END_IF

bRun_Auto:=TRUE;
//need to be set up an set point so the pump could keep the needed value in automatic mode
END_METHOD

METHOD INTERNAL m_CheckOper : BOOL
VAR_INPUT
END_VAR

VAR
	sMotorTypeAgrigate_to_check: STRING(2);
END_VAR
sMotorTypeAgrigate_to_check:=TO_STRING(Pump_ID);

IF sMotorTypeAgrigate_to_check='AG' THEN;
	m_CheckOper:=TRUE;
ELSE;
	IF stOperation.iActOperation=E_OperationButtons.ePlayAll THEN;
		m_CheckOper:=TRUE;
	ELSE;
		m_CheckOper:=FALSE;
	END_IF
END_IF
END_METHOD

METHOD m_Error : STRING(11)
VAR_INPUT
	
END_VAR
VAR
	skipTemp: BOOL;
END_VAR
//FB body not executed yet (first PLC cycle): Pump_ID and sID are not set
IF sID='' OR Pump_ID=E_Pump_List.eNotSelected THEN;
	RETURN;
END_IF

ton_RPM_feedback_lag_monitoring(PT:=T#10S);
IF __ISVALIDREF(stNidec) THEN;
	IF bRun
	AND ABS(stNidec.targetVelocity - nRPM_fdbk) > 10 
	THEN;
		ton_RPM_feedback_lag_monitoring.IN:=TRUE;
	ELSE;
		ton_RPM_feedback_lag_monitoring.IN:=FALSE;
	END_IF	
END_IF

CASE Pump_ID OF
	E_Pump_List.AG3001,
	E_Pump_List.AG3002,
	E_Pump_List.P3001,
	E_Pump_List.P3002,
	E_Pump_List.P1001,
	E_Pump_List.P4001,
	E_Pump_List.P4002,
	E_Pump_List.AG4001,
	E_Pump_List.AG4002,
	E_Pump_List.TB0001:;
		skipTemp:=TRUE;
ELSE;
		skipTemp:=FALSE;
END_CASE


IF bRun AND NOT skipTemp THEN;
	IF NOT DriveReady THEN;
		m_Error:=concat(sID,'x001');
		stOperation.bSetPause:=TRUE;
		RETURN;
	END_IF	

	IF ton_RPM_feedback_lag_monitoring.Q THEN;
		m_Error:=concat(sID,'x002');
		RETURN;
	END_IF
END_IF

IF NOT DriveReady AND NOT skipTemp THEN;
	m_Error:=concat(sID,'x003');
	//stOperation.bSetPause:=TRUE;
	RETURN;
END_IF


IF 	PressureSensor_ID <> E_ASense_Name.eNotSelected THEN;
	fbPressureSensor REF= fbAnalogSensor[PressureSensor_ID];
	IF __ISVALIDREF(fbPressureSensor) THEN;	
		ton_Pressure_feedback_monitoring(PT:=T#30S);
		IF bRun AND ( fbPressureSensor.bHH_Alarm 
					OR fbPressureSensor.bHH_Warning
					OR fbPressureSensor.bLL_Warning 
					OR fbPressureSensor.bLL_Alarm) 
		THEN;
			ton_Pressure_feedback_monitoring.IN:=TRUE;
		ELSE;
			ton_Pressure_feedback_monitoring.IN:=FALSE;
		END_IF	
		
		IF fbPressureSensor.bHH_Alarm AND ton_Pressure_feedback_monitoring.Q THEN;
			m_Error:=concat(sID,'x004');
			stOperation.bSetPause:=TRUE;
			RETURN;
		END_IF
		IF fbPressureSensor.bHH_Warning AND ton_Pressure_feedback_monitoring.Q THEN;
			m_Error:=concat(sID,'x005');
			RETURN;
		END_IF
		IF fbPressureSensor.bLL_Warning AND ton_Pressure_feedback_monitoring.Q THEN;
			m_Error:=concat(sID,'x006');
			RETURN;
		END_IF
		IF fbPressureSensor.bLL_Alarm AND ton_Pressure_feedback_monitoring.Q THEN;
			m_Error:=concat(sID,'x007');
			stOperation.bSetPause:=TRUE;
			RETURN;
		END_IF		
	END_IF	
END_IF

IF NOT modeAuto THEN;
	m_Error:=concat(sID,'x008');
	//stOperation.bSetPause:=TRUE;
	RETURN;
END_IF

m_Error:='';
END_METHOD

METHOD m_Get_Speed : INT
VAR_INPUT
END_VAR
m_Get_Speed:=nRPM_fdbk;
END_METHOD

METHOD m_Map_ControlWord : WORD
VAR_INPUT
	cwStruct : ControlWordStruct;
END_VAR
VAR
    tempWord : WORD;
END_VAR


// Map each bit from the structure to the corresponding bit in the control word
tempWord := 0;
IF cwStruct.SwitchOn THEN
    tempWord := tempWord OR 1; // Bit 0
END_IF
IF cwStruct.EnableVoltage THEN
    tempWord := tempWord OR 2; // Bit 1
END_IF
IF cwStruct.QuickStop THEN
    tempWord := tempWord OR 4; // Bit 2
END_IF
IF cwStruct.EnableOperation THEN
    tempWord := tempWord OR 8; // Bit 3
END_IF
// Reserved bits (4-7) are not set
IF cwStruct.FaultReset THEN
    tempWord := tempWord OR 256; // Bit 8
END_IF
// Reserved bits (9-15) are not set

m_Map_ControlWord := tempWord;
END_METHOD

METHOD m_Map_StatusWord : StatusWordStruct
VAR_INPUT
	wordInput : WORD;
END_VAR
VAR
    swStruct : StatusWordStruct;
END_VAR


// Map each bit from the status word to the corresponding field in the structure
swStruct.ReadyToSwitchOn    := (wordInput AND 1) <> 0;         // Bit 0
swStruct.SwitchedOn         := (wordInput AND 2) <> 0;         // Bit 1
swStruct.OperationEnabled   := (wordInput AND 4) <> 0;         // Bit 2
swStruct.Fault              := (wordInput AND 8) <> 0;         // Bit 3
swStruct.VoltageEnabled     := (wordInput AND 16) <> 0;        // Bit 4
swStruct.QuickStop          := (wordInput AND 32) <> 0;        // Bit 5
swStruct.SwitchOnDisabled   := (wordInput AND 64) <> 0;        // Bit 6
swStruct.Warning            := (wordInput AND 128) <> 0;       // Bit 7
swStruct.Remote             := (wordInput AND 256) <> 0;       // Bit 8
// Reserved bits (9-15) are not set, assuming FALSE
m_Map_StatusWord := swStruct;
END_METHOD

METHOD m_Nidec_Init : BOOL
VAR_INPUT
END_VAR
IF  NOT StatusWord.VoltageEnabled 
OR StatusWord.Fault 
OR (state_init=Ready AND NOT StatusWord.ReadyToSwitchOn )
THEN;
	ControlWord.SwitchOn:=FALSE;
	ControlWord.EnableVoltage:=FALSE;
	ControlWord.QuickStop:=FALSE;
	ControlWord.EnableOperation:=FALSE;
	ton_Drive_init(IN:=FALSE);
	state_init:=OFF;
	RETURN;
END_IF


CASE state_init OF
	OFF:; 
		IF TRUE
		AND StatusWord.VoltageEnabled
		AND StatusWord.QuickStop
		AND StatusWord.SwitchOnDisabled
		THEN;
			ton_Drive_init(IN:=TRUE,PT:=T#2S);
		ELSE;
			ton_Drive_init(IN:=FALSE);RETURN;
		END_IF
		
		IF ton_Drive_init.Q THEN;
			ControlWord.EnableVoltage:=TRUE;
			ControlWord.QuickStop:=TRUE;	
			state_init:=stage1;
			ton_Drive_init(IN:=FALSE);
		END_IF	
		
	stage1:;
		IF TRUE
		AND StatusWord.VoltageEnabled
		AND StatusWord.QuickStop
		AND NOT StatusWord.SwitchOnDisabled
		THEN;
			ton_Drive_init(IN:=TRUE,PT:=T#0.5S);
		ELSE;
			ton_Drive_init(IN:=FALSE);RETURN;
		END_IF
		
		IF ton_Drive_init.Q THEN;
			ControlWord.SwitchOn:=TRUE;
			state_init:=stage2;
			ton_Drive_init(IN:=FALSE);
		END_IF	
		
	stage2:;
		IF TRUE
		AND StatusWord.SwitchedOn
		AND StatusWord.VoltageEnabled
		AND StatusWord.QuickStop
		AND NOT StatusWord.SwitchOnDisabled
		THEN;
			ton_Drive_init(IN:=TRUE,PT:=T#0.5S);
		ELSE;
			ton_Drive_init(IN:=FALSE);RETURN;
		END_IF
		
		IF ton_Drive_init.Q THEN;
			state_init:=Ready;
			ton_Drive_init(IN:=FALSE);
		END_IF	

	
	
END_CASE
END_METHOD

METHOD m_Run : BOOL
VAR_INPUT
	RPM: REAL;
END_VAR
IF NOT bInitiated THEN;
	RETURN;
END_IF
bRun_Auto:=TRUE;
stPump.nRPM_Auto:=RPM;
m_Run:=TRUE;
END_METHOD

METHOD m_Stop : BOOL
VAR_INPUT
END_VAR
bRun_Auto:=FALSE;
bRun_Man:=FALSE;
m_Stop:=TRUE;
END_METHOD

END_FUNCTION_BLOCK

// ---- 00 Library/12 Analog Sensor/FB_AnalogSensor.TcPOU
FUNCTION_BLOCK FB_AnalogSensor
VAR_INPUT
	nSensorID	: 	E_ASense_Name	;
	nRawSensor	:	REAL				;
	arReset_AlrmWrn		:	ARRAY [0..3] OF BOOL		;//HH Alarm/LL Alarm/HH Warning/LL Warning
END_VAR
VAR_OUTPUT
	bLL_Alarm	:	BOOL	;
	bHH_Alarm	:	BOOL	;
	bLL_Warning	:	BOOL	;
	bHH_Warning	:	BOOL	;
END_VAR
VAR
	sName: STRING(12);

	stASens			:	REFERENCE TO ST_AnalogSensor	;
	state			: 	E_ASensor_State					;
	
	fbScaleFactor	: 	FB_ScaleFactor					;
	
	nTicks			:	INT:=0	;
	nI				:	INT		;
	
	bTestTemp		:	BOOL	;
	
	nTimeInCycles	:	INT:=100; //1 sec while cycletime is 10 ms
	nBufferSize_S	:	INT:=1	;//Buffer size in seconds
	nCycleTime_MS	:	INT:=10;//Cycle time in mili seconds
	
	
	//From Structure
	// Callibration 
	rawVal_Actual	: INT;//fb
	
	//MA
	arrRawVal_Actual	:	ARRAY [0..10000] OF INT	;//get out fb
	rTempRawVal			:	REAL	;//fb
	nRawSumm			:	DINT	;//fb
	
	bCopyRawTo_Min	: BOOL;//fb
	bCopyRawTo_Max	: BOOL;//fb
	
	//triggers
	arRS		:	ARRAY [0..3] OF RS		;//HH Alarm/LL Alarm/HH Warning/LL Warning
	
	ton_set_DATA: TON;
	rt_set_DATE: R_TRIG;
	fbScale: REFERENCE TO FB_ScaleFactor;
	fbMovingAverage: FB_MovingAverage;

	bSetFromTempCallibration: BOOL;
	bTypeTankConus: BOOL:=FALSE;
	rawTest: REAL;
END_VAR

nTimeInCycles:=TO_INT(nBufferSize_S*1000/nCycleTime_MS);
act_Get_Reference();
act_MA();
act_SetValues();
sName:=TO_STRING(nSensorID);
act_AlarmWarnings();

ACTION act_AlarmWarnings:
//arRS		:	ARRAY [0..3] OF RS		;//HH Alarm/LL Alarm/HH Warning/LL Warning
(*
arRS[0](
		SET:=(stASens.Value>= stASens.rHH_Alarm AND NOT bHH_Alarm) , 
		RESET1:=arReset_AlrmWrn[0] , Q1=>bHH_Alarm );
arRS[1](
		SET:=(stASens.Value<= stASens.rLL_Alarm AND NOT bLL_Alarm) , 
		RESET1:=arReset_AlrmWrn[1] , Q1=>bLL_Alarm );
arRS[2](
		SET:=(stASens.Value>= stASens.rHH_Warning AND stASens.Value<stASens.rHH_Alarm AND NOT bHH_Warning) , 
		RESET1:=arReset_AlrmWrn[2] , Q1=>bHH_Warning );
arRS[3](
		SET:=(stASens.Value<= stASens.rLL_Warning AND stASens.Value>stASens.rLL_Alarm AND NOT bLL_Warning) , 
		RESET1:=arReset_AlrmWrn[3] , Q1=>bLL_Warning );


*)		
bHH_Alarm:=stASens.Value>= stASens.rHH_Alarm;	
bLL_Alarm:=stASens.Value<= stASens.rLL_Alarm;	
bHH_Warning:=stASens.Value>= stASens.rHH_Warning AND stASens.Value<stASens.rHH_Alarm;	
bLL_Warning:=stASens.Value<= stASens.rLL_Warning AND stASens.Value>stASens.rLL_Alarm;
END_ACTION

ACTION act_Get_Reference:
stASens REF=g_AnalogSensor.stAnalogSensor[nSensorID];

stASens.ID:=TO_STRING(nSensorID);

//!!!!!!!!!!!!!!!!!!!!!!!!!!!!!!!!!!!!!!!!!!!!!!!!!!!!!!!!!!
//stASens.rawVal_Actual:=g_AnalogSensor.arAnalogSensorRawValue[nSensorID];
//stASens.rawVal_Actual:=nRawSensor;

//rTempRawVal:=rawTest;
CASE nSensorID OF 
	E_ASense_Name.LT3001,E_ASense_Name.LT3002,E_ASense_Name.LT4001,E_ASense_Name.LT4002:;
		bTypeTankConus:=TRUE;
ELSE;
		bTypeTankConus:=FALSE;
END_CASE
IF bTypeTankConus 
AND rTempRawVal<=stASens.rawVal_Min
THEN;
	stASens.Value:=mConus(rawValue:=rTempRawVal,baseIncriments:=stASens.rawVal_Min);
ELSE;
	fbScaleFactor(
		rVal:=rTempRawVal,//stASens.rawVal_Actual , 
		rInValHigh:=stASens.rawVal_Max , 
		rInValLow:=stASens.rawVal_Min , 
		rOutValHigh:=stASens.outVal_Max , 
		rOutValLow:=stASens.outVal_Min ,
		rOutOffset:=stASens.outOffset , 
		rValOut=>stASens.Value , 
		diValOut=>, 
		iValOut=> );	
END_IF

	
	
	
ton_set_DATA(PT:=T#20S, IN:=TRUE);
rt_set_DATE(CLK:=ton_set_DATA.Q);
IF rt_set_DATE.Q AND bSetFromTempCallibration THEN;
	set_Data(ID_reference:=nSensorID);
END_IF
END_ACTION

ACTION act_MA:
IF nTicks<nTimeInCycles THEN
	nTicks:=nTicks+1;
ELSIF nTicks>nTimeInCycles THEN
	nTicks:=nTimeInCycles;
END_IF

//moving ticks
nRawSumm:=0;
FOR nI:=nTimeInCycles TO 1 BY -1 DO
	arrRawVal_Actual[nI]:=arrRawVal_Actual[nI-1];
	//calculating summ
	nRawSumm:=nRawSumm+arrRawVal_Actual[nI];
END_FOR

arrRawVal_Actual[0]:=TO_INT(nRawSensor);
nRawSumm:=nRawSumm+arrRawVal_Actual[0];

rTempRawVal:=TO_REAL(nRawSumm/nTicks);


//fbMovingAverage(Value:=nRawSensor);
//rTempRawVal:=fbMovingAverage.Average;
END_ACTION

ACTION act_SetValues:
meth_SetRawValue(bSetValue:=bCopyRawTo_Max , nValToSet:=stASens.rawVal_Max , nRawValue:=rawVal_Actual );
meth_SetRawValue(bSetValue:=bCopyRawTo_Min , nValToSet:=stASens.rawVal_Min , nRawValue:=rawVal_Actual );
END_ACTION

METHOD mConus : REAL
VAR_INPUT
	rawValue: REAL;
	baseIncriments: REAL;
END_VAR



VAR
	hFactor: REAL;
	baseIncriment: REAL := 1050;
	h: REAL := 140;
	ConusConstant: REAL := 0.00000002165;
	pi: REAL:=3.1415926535;
	k: REAL:=3000000; // convert mm^3 to liters


	radius: REAL := 525;
	vConus: REAL;
END_VAR

VAR
	
END_VAR


//hFactor:=baseIncriment*h;

vConus:=pi*radius*radius*h/k;
IF baseIncriments=0 THEN;
	RETURN;
END_IF
ConusConstant:=vConus/(baseIncriments * baseIncriments * baseIncriments);
mConus:=ConusConstant*rawValue*rawValue*rawValue;
END_METHOD

METHOD INTERNAL meth_SetRawValue : BOOL
VAR_IN_OUT
	bSetValue	:	BOOL	;
	nValToSet	:	REAL	;
END_VAR
VAR_INPUT
	nRawValue	:	REAL		;
END_VAR
IF bSetValue THEN
	nValToSet:=nRawValue;
	bSetValue:=FALSE;
END_IF
END_METHOD

METHOD mSetAsConus : BOOL
VAR_INPUT
END_VAR
bTypeTankConus:=TRUE;
END_METHOD

METHOD set_Data : BOOL
VAR_INPUT
	ID_reference: E_ASense_Name;
END_VAR
fbScale REF= gIO.fbScaleFactor[ID_reference];
IF NOT __ISVALIDREF(fbScale) THEN;
	RETURN;
END_IF
	


stASens.rawVal_Max:=fbScale.rInValHigh;
stASens.rawVal_Min:=fbScale.rInValLow;
stASens.outVal_Max:=fbScale.rOutValHigh;
stASens.outVal_Min:=fbScale.rOutValLow;
stASens.outOffset:=fbScale.rOutOffset;
END_METHOD

END_FUNCTION_BLOCK

// ---- 00 Library/30 IO/FB_ScaleFactor.TcPOU
FUNCTION_BLOCK FB_ScaleFactor
VAR_INPUT
	rVal: REAL;
	rInValHigh: REAL;
	rInValLow: REAL;
	rOutValHigh: REAL;
	rOutValLow: REAL;
	rOutOffset: REAL:=0;
END_VAR

VAR
	rOfset: REAL;
	a: REAL;
	b: REAL;
END_VAR
VAR_OUTPUT
	rValOut: REAL;
	diValOut: DINT;
	iValOut: INT;
END_VAR

IF rInValHigh-rInValLow<>0 THEN;
	a:=(rOutValHigh-rOutValLow)/(rInValHigh-rInValLow);
ELSE;
	a:=0;
END_IF
b:=rOutValHigh-(a*rInValHigh);
rValOut:=(a*rVal+b)+rOutOffset;
diValOut:=TRUNC(rValOut);
iValOut:=DINT_TO_INT(diValOut);

END_FUNCTION_BLOCK

// ---- 00 Library/10 Utils/FB_MovingAverage.TcPOU
FUNCTION_BLOCK FB_MovingAverage
VAR_INPUT
	Value: REAL;
END_VAR
VAR_OUTPUT
	Average: REAL;

END_VAR
VAR
	arr: ARRAY[1..cMaxBufer] OF REAL;

	Sum: REAL;
	i: INT;
END_VAR
VAR CONSTANT
	cMaxBufer: INT:=500; // 10msec * 500 = 5 sec

END_VAR

Sum:=0;
FOR	i:=1 TO cMaxBufer DO
	Sum:=Sum+arr[i];
END_FOR


Average:=Sum/cMaxBufer;
FOR i:=cMaxBufer TO 2 BY-1 DO
	arr[i]:=arr[i-1];
END_FOR
arr[1]:=Value;

END_FUNCTION_BLOCK

// ---- 00 Library/02 Pump/02.1 Dosing Pump/FB_DosingPump.TcPOU
FUNCTION_BLOCK FB_DosingPump EXTENDS FB_SFC_Cycle
VAR_INPUT
END_VAR
VAR_OUTPUT
	valve_A			: BOOL;
	valve_B			: BOOL;
END_VAR
VAR

	action_Time		: TIME:=T#0.5S;
	startDelay		: TIME:=T#0S;
	
	reqTiks			: DINT:=5;
	actTiks			: DINT:=5;
	
	fStageVolume	: REAL:=65; 	// CC/stage
	fReqVolume		: REAL:=500.0; 	// CC
	fActVolume		: REAL; 		// CC


END_VAR

VAR PERSISTENT
	
END_VAR

act_GetReference();

act_Oper();

reqTiks:=TRUNC(fReqVolume/fStageVolume);
fActVolume:=(actTiks*fStageVolume);

ACTION _acheck_Count_active:
bStepDone:=FALSE;
IF actTiks>=reqTiks THEN;
	bStepDone:=TRUE;
END_IF
END_ACTION

ACTION _acheck_Count_entry:
actTiks:=actTiks+1;
END_ACTION

ACTION _aDone_entry:
bRun:=FALSE;
bDone:=TRUE;
END_ACTION

ACTION _aInit_act_Oper_active:
SFCReset:=FALSE;
END_ACTION

ACTION _aInit_act_Oper_exit:
valve_A:=valve_B:=bRun:=bDone:=FALSE;
END_ACTION

ACTION _aReady_exit:
actTiks:=0;
END_ACTION

ACTION _astage_A_entry:
valve_A:=TRUE;
END_ACTION

ACTION _astage_A_exit:
valve_A:=FALSE;
END_ACTION

ACTION _astage_B_entry:
valve_B:=TRUE;
END_ACTION

ACTION _astage_B_exit:
valve_B:=FALSE;
END_ACTION

ACTION act_GetReference:
m_Set_SFCFlags_Reference();
END_ACTION

ACTION act_Oper:
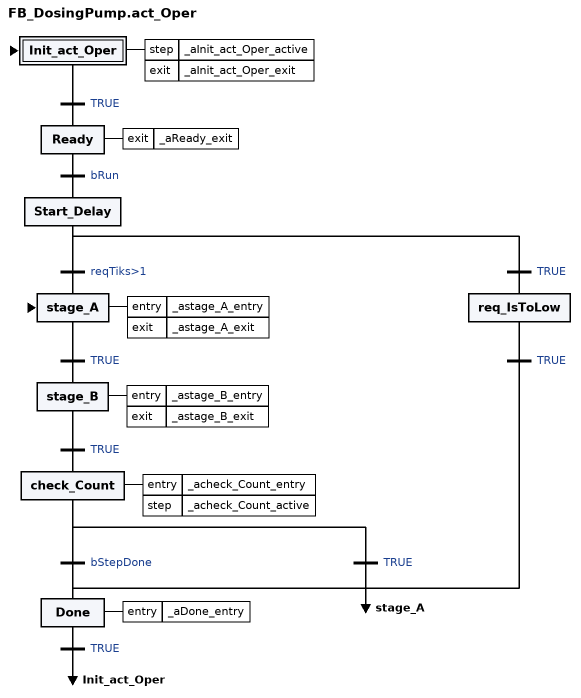
INITIAL_STEP Init_act_Oper:
    _aInit_act_Oper_active(N);  // step action
    _aInit_act_Oper_exit(P0);  // exit action
END_STEP
TRANSITION FROM Init_act_Oper TO Ready
    := TRUE;
END_TRANSITION
STEP Ready:
    _aReady_exit(P0);  // exit action
END_STEP
TRANSITION FROM Ready TO Start_Delay
    := bRun;
END_TRANSITION
STEP Start_Delay:  // min time startDelay
END_STEP
TRANSITION FROM Start_Delay TO stage_A
    := reqTiks>1;
END_TRANSITION
STEP stage_A:  // min time action_Time
    _astage_A_entry(P1);  // entry action
    _astage_A_exit(P0);  // exit action
END_STEP
TRANSITION FROM stage_A TO stage_B
    := TRUE;
END_TRANSITION
STEP stage_B:  // min time action_Time
    _astage_B_entry(P1);  // entry action
    _astage_B_exit(P0);  // exit action
END_STEP
TRANSITION FROM stage_B TO check_Count
    := TRUE;
END_TRANSITION
STEP check_Count:
    _acheck_Count_entry(P1);  // entry action
    _acheck_Count_active(N);  // step action
END_STEP
TRANSITION FROM check_Count TO Done
    := bStepDone;
END_TRANSITION
TRANSITION FROM check_Count TO stage_A
    := TRUE;
END_TRANSITION
TRANSITION FROM Start_Delay TO req_IsToLow
    := TRUE;
END_TRANSITION
STEP req_IsToLow:
END_STEP
TRANSITION FROM req_IsToLow TO Done
    := TRUE;
END_TRANSITION
STEP Done:
    _aDone_entry(P1);  // entry action
END_STEP
TRANSITION FROM Done TO Init_act_Oper
    := TRUE;
END_TRANSITION
// branch label Branch0_act_Oper
// branch label Branch1_act_Oper
END_ACTION

METHOD m_RunVolume : BOOL
VAR_INPUT
	Volume	:REAL;
END_VAR
fReqVolume:=Volume;
mRun();
IF rtDone.Q THEN;
	m_RunVolume:=TRUE;	
END_IF
END_METHOD

METHOD m_Set_SFCFlags_Reference : BOOL
//Set reference to SFC flags

refSFC.SFCInit REF= SFCInit;
refSFC.SFCReset REF= SFCReset;
refSFC.SFCError REF= SFCError;
refSFC.SFCEnableLimit REF= SFCEnableLimit;
refSFC.SFCErrorStep REF= SFCErrorStep;
refSFC.SFCErrorPOU REF= SFCErrorPOU;
refSFC.SFCQuitError REF= SFCQuitError;
refSFC.SFCPause REF= SFCPause;
refSFC.SFCTrans REF= SFCTrans;
refSFC.SFCCurrentStep REF= SFCCurrentStep;
refSFC.SFCTip REF= SFCTip;
refSFC.SFCTipMode REF= SFCTipMode;

// Cycle handle for SFC
m_SFC_Handle();
END_METHOD

METHOD m_Stop : BOOL
VAR_INPUT
END_VAR
SFCReset:=TRUE;
END_METHOD

END_FUNCTION_BLOCK

// ---- 00 Library/HeatExchenger/FB_HeatExchanger.TcPOU
FUNCTION_BLOCK FB_HeatExchanger
VAR_IN_OUT
	stHeatExchanger	:	ST_HeatExchanger	;
END_VAR
VAR_INPUT
	nValveID		:	E_Pis_Name 	;	
	nAnalogValveID	:	E_Pis_Name 	;

	nProcCntrlID	:	E_ProcessControl_Name	;
END_VAR
VAR_OUTPUT
	nAlagonValveCntrOut	:	INT	;//output for analog valve opening
END_VAR
VAR
	stPis			:	REFERENCE TO ST_Piston;
	stPisAnalog		:	REFERENCE TO ST_Piston;
	
	stProcessControl		:	REFERENCE TO ST_ProcessControl	;
	fbProcessControl		: 	REFERENCE TO FB_ProcessControl	;
END_VAR

act_GetReference();
//act_AnalogOutScaling();

stProcessControl.fCtrlOutput_Min:=0;
stProcessControl.fCtrlOutput_Max:=100;
stProcessControl.rValue_Min_To_ReleaseControl:=15; //Degrees

//PID MANUAL follows HMI request in any CIP state; in manual PID output = stProcessControl.fCtrlOutput_Manual (from HMI)
fbProcessControl.mManual(value:=stHeatExchanger.bManual);
//Automatic: PID held in reset while control is not active (output 0, every start begins from 0)
stProcessControl.bReset:=NOT stHeatExchanger.bManual AND NOT stProcessControl.bActiveCntr;

//On-Off valve is controlled only in automatic
IF NOT stHeatExchanger.bManual THEN;
	IF stProcessControl.bActiveCntr AND NOT stPis.st_Open THEN
		stPis.req_Open:=TRUE;
	ELSIF NOT stProcessControl.bActiveCntr AND NOT stPis.st_Close THEN
		stPis.req_Close:=TRUE;
	END_IF
	
END_IF
//Manual: output directly from HMI value (PID stays in MANUAL for bumpless return to automatic)
IF stHeatExchanger.bManual THEN;
	nAlagonValveCntrOut:=mCMD_to_Analog(fControl:=LIMIT(stProcessControl.fCtrlOutput_Min, stProcessControl.fCtrlOutput_Manual, stProcessControl.fCtrlOutput_Max));
ELSIF stProcessControl.bActiveCntr THEN;
	nAlagonValveCntrOut:=mCMD_to_Analog(fControl:=stProcessControl.fCtrlOutput);
ELSE;
	//Control not active: analog valve closed, V1032 closes
	nAlagonValveCntrOut:=0;
END_IF
IF nAlagonValveCntrOut=0 AND NOT stPisAnalog.st_Close THEN;
	stPisAnalog.req_Close:=TRUE;
ELSIF nAlagonValveCntrOut<>0 AND NOT stPisAnalog.st_Open THEN;
	stPisAnalog.req_Open:=TRUE;
END_IF

ACTION act_AnalogOutScaling:
IF (stHeatExchanger.cntrlVal_Max-stHeatExchanger.cntrlVal_Min)<>0 THEN
	nAlagonValveCntrOut:=DINT_TO_INT((TRUNC((stProcessControl.fCtrlOutput*
		(stHeatExchanger.outVal_Max-stHeatExchanger.outVal_Min)/(stHeatExchanger.cntrlVal_Max-stHeatExchanger.cntrlVal_Min))+
		stHeatExchanger.outOffset)));
END_IF
END_ACTION

ACTION act_GetReference:
//On-Off walve structure
stPis REF= g_Piston.stPis[nValveID];
stPisAnalog REF= g_Piston.stPis[nAnalogValveID];

stProcessControl REF=g_ProcControl.arr_stProcCntrl[nProcCntrlID];
fbProcessControl REF=g_ProcControl.arr_fbProcCntrl[nProcCntrlID];
END_ACTION

METHOD m_Auto : BOOL
VAR_INPUT
END_VAR
END_METHOD

METHOD m_Run : BOOL
VAR_INPUT
END_VAR
END_METHOD

METHOD m_Stop : BOOL
VAR_INPUT
END_VAR
END_METHOD

METHOD mCMD_to_Analog : INT
VAR_INPUT
	fControl: LREAL;
END_VAR
IF (stHeatExchanger.cntrlVal_Max-stHeatExchanger.cntrlVal_Min)<>0 THEN
	mCMD_to_Analog:=DINT_TO_INT((TRUNC((fControl*
		(stHeatExchanger.outVal_Max-stHeatExchanger.outVal_Min)/(stHeatExchanger.cntrlVal_Max-stHeatExchanger.cntrlVal_Min))+
		stHeatExchanger.outOffset)));
ELSE;
	mCMD_to_Analog:=0;
END_IF

//nAlagonValveCntrOut
END_METHOD

END_FUNCTION_BLOCK

// ---- 00 Library/Sensors/FB_TankSensors.TcPOU
FUNCTION_BLOCK FB_TankSensors
VAR_IN_OUT
	stTankLevel	:	ST_Tank_Level	;
END_VAR
VAR_INPUT
	volume: REAL:=100; //litr
	//Level
	senHL				:	BOOL	;
	senLL				:	BOOL	;
	nSensorLvl_ID		: 	E_ASense_Name	;
	nSensorLvl_Raw		:	INT		;
	//Temperature
	nSensorTemp_ID		: 	E_ASense_Name	;
	nSensorTemp_Raw		:	INT		;
END_VAR
VAR_OUTPUT
	act_Volume			: REAL;
END_VAR
VAR
	stASensLvl			:	REFERENCE TO ST_AnalogSensor	;
	
	stASensTemp			:	REFERENCE TO ST_AnalogSensor	;
	
	Call_TankLevel			:	FB_AnalogSensor	;
	Call_TankTemp			:	FB_AnalogSensor	;
	tonEmpty: TON;
END_VAR

//Call_TankLevel(nSensorID:=nSensorLvl_ID, nRawSensor:=nSensorLvl_Raw );
//Call_TankTemp(nSensorID:=nSensorTemp_ID, nRawSensor:=nSensorTemp_Raw );
act_TankLvl();
act_Volume:=stTankLevel.rTankLevel;

ACTION act_TankLvl:
stASensLvl REF=g_AnalogSensor.stAnalogSensor[nSensorLvl_ID];

IF stTankLevel.bIn_LL_signal=FALSE AND stTankLevel.bIn_HL_signal=FALSE THEN
	tonEmpty.IN:=TRUE;
ELSE;
	tonEmpty.IN:=FALSE;
END_IF
IF stTankLevel.bIn_LL_signal=TRUE AND stTankLevel.bIn_HL_signal=FALSE THEN
	stTankLevel.e_state:=E_Tank_Level.eLL;
ELSIF stTankLevel.bIn_LL_signal=TRUE AND stTankLevel.bIn_HL_signal=TRUE THEN
	stTankLevel.e_state:=E_Tank_Level.eHL;
ELSIF stTankLevel.bIn_LL_signal=FALSE AND stTankLevel.bIn_HL_signal=TRUE THEN
	stTankLevel.e_state:=E_Tank_Level.eERROR;
END_IF

stTankLevel.rTankLevel:=stASensLvl.Value;
stTankLevel.rTankLevelPercentage:=stTankLevel.rTankLevel/volume*100;
stTankLevel.bIn_HL_signal:=senHL;
stTankLevel.bIn_LL_signal:=senLL;

tonEmpty(PT:=T#3S);
IF tonEmpty.Q THEN;
	stTankLevel.e_state:=E_Tank_Level.eEmpty;
END_IF
END_ACTION

